(* IEC 61131-3 sources: daoli-st-library/DL_MathData (part 18) *)

(* ---- FC_DL_LrealToFixedField.st ---- *)
(*==============================================================================
 * 组件名称 (Component)  : FC_DL_LrealToFixedField
 * 溯源说明 (Provenance): 道莅 clean-room 防御性实现（IEC 61131-3 纯净实现，闭源文档仅借语义，零代码行）
 * 所属子库 (Sublibrary) : DL_MathData / DataFormat
 * 当前版本 (Version)    : 1.0.0
 * 兼容性   (Platform)   : CODESYS 3.5 / TwinCAT 3 / 汇川 InoProShop / 施耐德
 *                         Machine Expert；纯 IEC 61131-3（第 3 版），仅用
 *                         Standard.library 的 MID / CONCAT / LEN / ABS / TRUNC / LIMIT
 * 组件分类 (Category)   : 函数（FUNCTION）· 纯函数 · 浮点 → 定宽定点文本
 * 功能一句话 (Summary)  : 把 LREAL 按指定整数位宽与小数位数输出成定宽定点文本
 *                         （四舍五入或截断、可选强制正号），非有限输入拒绝输出。
 *
 * 【填充与对齐规则（与 FC_DL_IntToFixedField 共用同一段口径原文）】
 *   ① 右对齐：数值永远贴字段右端，填充字符只在左侧。
 *   ② 本件无 bZeroPad 引脚，整数部分统一用**空格**填充到 uIntDigits 位
 *      ——即 #1 的 bZeroPad = FALSE 分支口径；领先零一律压成空格，
 *      但至少保留一位数字（0.5 输出 "0.500" 而非 ".500"）。
 *   ③ 符号位占一位：**恒留一格**（无符号时填空格），故字段总宽恒为
 *      1 + uIntDigits + (uDecDigits > 0 ? 1 + uDecDigits : 0) ≤ 23，
 *      定长报文的列位由此确定，不随数值正负漂移。
 *   ④ 宽度是契约：uIntDigits / uDecDigits 越界只钳位（0460 信息级）；
 *      整数部分装不下时不截断，直接饱和到全 9 并置 bSaturated。
 *
 * 本件存在的意义 (Why this unit exists)
 *   MES 称重/流量报文要的是「固定小数位、列位对齐」的数值域（"  1234.567"）。
 *   平台内建 LREAL_TO_STRING 的小数位口径与科学计数法门槛三平台不一致
 *   （CODESYS / TwinCAT / InoProShop 对同一值可能给出不同尾数与指数形式），
 *   故本件**禁用** LREAL_TO_STRING，自行按 10 的幂分解：绝对值域取整 → 逐位
 *   分解 → 拼接，末位再加符号，天然对称，输出可在三平台逐字节比对。
 *
 * 边界安全 (Boundary)
 *   ① 非有限输入：NaN 用自不等判据 (x−x) <>(x−x)，±Inf 用 ABS(x) > DBL_MAX
 *      精确判据（R79，禁近似阈值）→ 故障 03AE、bValid = FALSE，
 *      **绝不输出 'NaN' / 'Inf' 冒充合法报文**；
 *   ② uIntDigits 钳 1~15、uDecDigits 钳 0~6，越界钳位 + 信息 0460；
 *   ③ 字段装不下（1 + 整数位 + 1 + 小数位 > 24）→ 故障 03AF。钳位后最大为
 *      23，本分支结构性不可达，属纯防御纵深（R94 统一后处理）；
 *   ④ 整数部分有效位超 uIntDigits → 饱和全 9 + bSaturated + 信息 0461，
 *      bValid 保持 TRUE（饱和可观测，与「非有限」性质不同）；
 *   ⑤ 四舍五入实际进位导致整数位溢出 → 同一饱和路径（复用 0461，不新开码，R90）；
 *   ⑥ 舍入进位未溢出整数位 → 信息 0460 复用（R90 不加码，头注释写明复用理由）；
 *   ⑦ 全部取整只用 TRUNC 作用于**小于 10 的商与小于 10^d 的余数**，绝不 TRUNC
 *      大数，因此任何平台都不会在内建转换上溢出。
 * 遗留假设 (Assumption)
 *   整数部分超过 15 位十进制时 LREAL 已无精确表示（2^53 ≈ 9.007E15），
 *   本件按「输入本身已失真」处理，不承诺末位准确；这也是把
 *   uIntDigits 上限定为 15 的原因（DL_FF_INTMAX）。
 *   逐位分解的商与余数为浮点运算，末位可能受二进制表示误差影响 ±1 个最小
 *   单位（已在四舍五入阈值中吸收），不承诺与十进制手算逐位一致。
 *
 * 错误码    : 16#0001_0460 整数位/小数位已钳位，或四舍五入发生进位——信息级，正常防御
 *             16#0001_0461 整数部分有效位超出字段宽度，已饱和为全 9——信息级，饱和可观测
 *             16#0001_03AE 输入非有限（NaN / ±Inf），拒绝输出——故障级，返回 FALSE
 *             16#0001_03AF 字段宽度装不下（整数位+小数位+符号+小数点超上限）——故障级
 *             16#0001_03B0 预留禁用（故障级，不得挪用）
 * 码位总账  : 16#0001_0460 用 / 16#0001_0461 用 ｜ 16#0001_03AE 用 / 16#0001_03AF 用 / 16#0001_03B0 预留
 * 状态机    : N/A —— 纯函数无顺序状态机
 * 采样约定  : 纯组合函数，无定时器、无内部驻留状态
 * 依赖说明  : 无 DL_ 内部依赖；仅 Standard.library 的 MID / CONCAT / LEN / ABS / TRUNC / LIMIT
 * 验收向量  : V1 1234.5678/整数6/小数3/四舍五入 → '  1234.568'，写 11，TRUE
 *             V2 -42.5/整数6/小数3/截断 → '   -42.500'，写 11，TRUE
 *             V3 0.5/整数2/小数2 → '  0.50'，写 6，TRUE（领先零压成空格但保留一位）
 *             V4 999999.9999/整数6/小数3/四舍五入 → 饱和全 9 ' 999999.999'，
 *                bSaturated=TRUE，eErr=0461，TRUE（进位溢出主向量）
 *             V5 NaN → FALSE，sField=''，eErr=03AE，bError=TRUE
 *             V6 +Inf → FALSE，eErr=03AE
 *             V7 整数位 0 / 小数位 9 → 钳到 1 / 6 且 eErr=0460，仍返回 TRUE
 *             V8 1.0E16/整数15/小数0 → 饱和全 9（失真声明主向量）
 * 红线自检  : 全局变量声明零使用 / 外部变量访问零使用 / 物理地址零使用 ｜ 纯 IEC 61131-3（零厂商转换）
 *             浮点无判等比较（仅自不等 NaN 判据与容差阈值）｜ 除法前置判零
 *             （fPow 恒 ≥ 1.0，构造性非零）｜ 循环全部带守卫 ｜ 数组下标前置界检
 *             全变量双语同行注释 ｜ 状态机 N/A ｜ 无定时器实例 ｜ 无魔法数
 * 修订历史  : 2026-11-16  v1.0.0  首版入库（R22 · 批 1 · 定宽数值字段族）
 *============================================================================*)

FUNCTION FC_DL_LrealToFixedField : BOOL
VAR_INPUT
    fValue      : LREAL;                       // 待编码浮点值，任意有限值 / value to encode, any finite value
    uIntDigits  : UINT := 6;                   // 整数部分最少字符数 [字符]，范围 1~15 / minimum integer characters, range 1~15
    uDecDigits  : UINT := 3;                   // 小数位数 [位]，范围 0~6 / decimal digits, range 0~6
    bRound      : BOOL := TRUE;                // TRUE 四舍五入 / FALSE 向零截断 / TRUE rounds half up, FALSE truncates
    bForceSign  : BOOL := FALSE;               // 正数是否强制 '+' 号 / force '+' sign on positive values
END_VAR
VAR_OUTPUT
    sField      : STRING(24);                  // 定宽定点文本，右对齐 [ASCII] / fixed width fixed point text, right aligned
    uFieldLen   : UINT;                        // 实际写入字符数 [字符] / actual written length [char]
    bSaturated  : BOOL;                        // 整数部分已饱和为全 9 / integer part saturated to all nines
    eErr        : UDINT;                       // 错误码，0 表示无错 / error code, 0 means no error
    bError      : BOOL;                        // 故障级标志，仅故障级错误置位 / fault-class flag, set only on fault-level codes
    bValid      : BOOL;                        // 结果可用标志（饱和时仍为 TRUE） / result usable flag, still TRUE when saturated
END_VAR
VAR
    nIntUse     : INT;                         // 生效整数位宽 [字符]，已钳位 1~15 / effective integer width, clamped
    nDecUse     : INT;                         // 生效小数位数 [位]，已钳位 0~6 / effective decimal digits, clamped
    nTotal      : INT;                         // 字段总宽 [字符] / total field width
    nLead       : INT;                         // 首个非零整数位下标 [索引]，0 表示全零 / index of the first non-zero integer digit, 0 when all zero
    nI          : INT;                         // 通用循环下标 [索引] / general loop index
    nJ          : INT;                         // 升序循环变量（镜像下标用）[索引] / ascending loop var for mirrored index
    nGuard      : INT;                         // 循环守卫计数器 [次] / loop guard counter
    nFracMax    : LINT;                        // 小数位满量 10^nDecUse [无量纲] / full range of the decimal part
    liFrac      : LINT;                        // 小数部分放大后的整数值 [无量纲] / scaled integer value of the decimal part
    liDig       : LINT;                        // 单步取位结果 [无量纲] / single digit extraction result
    bNeg        : BOOL;                        // 输入为负 / input is negative
    bNeedSign   : BOOL;                        // 是否输出符号字符 / whether a sign character is emitted
    bAllNine    : BOOL;                        // 饱和全 9 路径 / saturated all-nines path
    bCarry      : BOOL;                        // 舍入发生进位 / rounding produced a carry
    bPropagate  : BOOL;                        // 进位仍在传播 / the carry is still propagating
    fAbs        : LREAL;                       // 输入绝对值 [无量纲] / absolute value of the input
    fRem        : LREAL;                       // 未分解的剩余量 [无量纲] / remaining undecomposed value
    fPow        : LREAL;                       // 当前位的 10 的幂 [无量纲] / power of ten of the current position
    fIntLimit   : LREAL;                       // 整数部分容量 10^nIntUse [无量纲] / integer capacity
    fFracScaled : LREAL;                       // 放大后的小数部分 [无量纲] / scaled decimal part
    fDiff       : LREAL;                       // NaN 自不等判据的中间量 [无量纲] / intermediate for the NaN self-inequality test
    aInt        : ARRAY[1..15] OF USINT;       // 整数位数字缓存，1 基 [无量纲] / integer digit cache, 1-based
    aDec        : ARRAY[1..6] OF USINT;        // 小数位数字缓存，1 基 [无量纲] / decimal digit cache, 1-based
    sInt        : STRING(15);                  // 整数段（含空格填充）[ASCII] / integer segment including space padding
    sFrac       : STRING(6);                   // 小数段 [ASCII] / decimal segment
    sSign       : STRING(1);                   // 符号段，无符号时填空格 [ASCII] / sign segment, a space when unsigned
    sDigitCh    : STRING(1);                   // 单字符数字，由数字表取出 [ASCII] / single digit character taken from the table
END_VAR
VAR CONSTANT
    DL_FF_MAXLEN   : UINT := 24;               // STRING(24) 物理上限 [字符]，禁写成 255 / physical bound of STRING(24), never 255
    DL_FF_INTMAX   : UINT := 15;               // 整数位宽上限 [字符]，受 2^53 精度约束 / integer width ceiling, bounded by 2^53
    DL_FF_DECMAX   : UINT := 6;                // 小数位数上限 [位] / decimal digit ceiling
    DL_FF_MAXLEN_I : INT := 24;                // 字段上限的 INT 副本 [字符] / INT copy of the field ceiling
    DL_INT_MIN     : INT := 1;                 // 整数位宽下限 [字符] / integer width floor
    DL_DEC_MIN     : INT := 0;                 // 小数位数下限 [位] / decimal digit floor
    DL_INT_MAX     : INT := 15;                // 整数位宽上限的 INT 副本 [字符] / INT copy of the integer width ceiling
    DL_DEC_MAX     : INT := 6;                 // 小数位数上限的 INT 副本 [位] / INT copy of the decimal digit ceiling
    DL_U_ZERO      : UINT := 0;                // 无符号零值 [无量纲] / unsigned zero
    DL_U_ONE       : UINT := 1;                // 无符号一值 [无量纲] / unsigned one
    DL_ONE_I       : INT := 1;                 // 整型一，用于 FOR 起始 [无量纲] / integer one used as a FOR start
    DL_SIGN_RES    : INT := 1;                 // 符号位恒留宽度 [字符] / reserved sign position width
    DL_POINT_W     : INT := 1;                 // 小数点占位宽度 [字符] / decimal point width
    DL_DIG_LAST    : INT := 9;                 // 单个数字位最大值 [无量纲] / maximum single digit value
    DL_GUARD_MAX   : INT := 20;                // 循环守卫上限 [次] / loop guard ceiling
    DL_TEN_I       : INT := 10;                // 十进制基数的 INT 副本 [无量纲] / INT copy of the decimal radix
    DL_TEN_L       : LINT := 10;               // 十进制基数的 LINT 副本 [无量纲] / LINT copy of the decimal radix
    DL_TEN_R       : LREAL := 10.0;            // 十进制基数的 LREAL 副本 [无量纲] / LREAL copy of the decimal radix
    DL_ONE_R       : LREAL := 1.0;             // 实型一，幂循环起点 [无量纲] / real one, power loop start
    DL_HALF_R      : LREAL := 0.5;             // 四舍五入偏置 [无量纲] / half-up rounding offset
    DL_LREAL_MAX   : LREAL := 1.7976931348623157E308; // LREAL 最大有限值，±Inf 精确判据 / maximum finite LREAL, exact infinity test
    DL_DIGITS      : STRING(10) := '0123456789'; // 数字字符表，经 MID 取值 [ASCII] / digit table read through MID
    DL_POINT_CH    : STRING(1) := '.';         // 小数点字符 [字符] / decimal point character
    DL_SPACE_CH    : STRING(1) := ' ';         // 空格填充字符 [字符] / space pad character
    DL_SIGN_PLUS   : STRING(1) := '+';         // 正号字符 [字符] / plus sign character
    DL_SIGN_MINUS  : STRING(1) := '-';         // 负号字符 [字符] / minus sign character
    DL_CH_ONE      : INT := 1;                 // MID 的单字符长度 [字符] / single character length for MID
END_VAR

(*------------------------------------------------------------------------------
 * 段 1｜返回值与输出预置（L1/L9：任何早退路径不留脏值）
 *      Preset the return value and every output, no stale value on any exit
 *-----------------------------------------------------------------------------*)
FC_DL_LrealToFixedField := FALSE;              // 返回值预置失败 / preset to FALSE
sField      := '';                             // 字段清空 / field cleared
uFieldLen   := 0;                              // 写入长度预置 0 [字符] / written length preset to zero
bSaturated  := FALSE;                          // 饱和标志预置 FALSE / saturation preset to FALSE
eErr        := 16#0000_0000;                   // 错误码预置无错 / error code preset to none
bError      := FALSE;                          // 故障标志预置 FALSE / fault flag preset to FALSE
bValid      := FALSE;                          // 结果可用预置 FALSE / usable flag preset to FALSE
nIntUse     := DL_INT_MIN;                     // 整数位宽预置下限 / integer width preset to the floor
nDecUse     := DL_DEC_MIN;                     // 小数位数预置下限 / decimal digits preset to the floor
nTotal      := 0;                              // 总宽预置 0 / total width preset to zero
nLead       := 0;                              // 领先零位置预置 0 / leading position preset to zero
nGuard      := 0;                              // 守卫预置 0 / guard preset to zero
nFracMax    := 1;                              // 小数满量预置 1 / decimal full range preset to one
liFrac      := 0;                              // 小数整数化预置 0 / scaled decimal preset to zero
liDig       := 0;                              // 取位结果预置 0 / digit result preset to zero
bNeg        := FALSE;                          // 负号标志预置 FALSE / negative flag preset to FALSE
bNeedSign   := FALSE;                          // 符号标志预置 FALSE / sign flag preset to FALSE
bAllNine    := FALSE;                          // 饱和路径预置 FALSE / saturation path preset to FALSE
bCarry      := FALSE;                          // 进位标志预置 FALSE / carry flag preset to FALSE
bPropagate  := FALSE;                          // 进位传播预置 FALSE / propagation preset to FALSE
fAbs        := 0.0;                            // 绝对值预置 0 / absolute value preset to zero
fRem        := 0.0;                            // 剩余量预置 0 / remainder preset to zero
fPow        := DL_ONE_R;                       // 幂预置 1 / power preset to one
fIntLimit   := DL_ONE_R;                       // 整数容量预置 1 / integer capacity preset to one
fFracScaled := 0.0;                            // 放大值预置 0 / scaled value preset to zero
sSign       := DL_SPACE_CH;                    // 符号段预置空格（符号位恒留一格） / sign segment preset to a space, the position is always reserved

(*------------------------------------------------------------------------------
 * 段 2｜非有限输入闸门（R79 精确判据：NaN 自不等 + ±Inf 与 DBL_MAX 直比）
 *      Non-finite gate with exact criteria, no approximate thresholds
 *-----------------------------------------------------------------------------*)
fDiff := fValue - fValue;                      // 有限值得 0，NaN 得 NaN / zero for finite input, NaN for NaN input
IF fDiff <> fDiff THEN
    eErr   := 16#0001_03AE;                    // 故障级：NaN 输入 / fault: NaN input
    bError := TRUE;                            // 置故障标志 / raise the fault flag
    bValid := FALSE;                           // 结果不可用 / result unusable
    sField := '';                              // 绝不输出 'NaN' 冒充合法报文 / never emit NaN as a legal field
    RETURN;                                    // 早退路径已统一后处理 / the early exit is fully post-processed
END_IF
IF ABS(fValue) > DL_LREAL_MAX THEN
    eErr   := 16#0001_03AE;                    // 故障级：±Inf 输入 / fault: infinity input
    bError := TRUE;                            // 置故障标志 / raise the fault flag
    bValid := FALSE;                           // 结果不可用 / result unusable
    sField := '';                              // 绝不输出 'Inf' 冒充合法报文 / never emit Inf as a legal field
    RETURN;
END_IF

(*------------------------------------------------------------------------------
 * 段 3｜位宽钳位（越界只钳位；信息级码不置 bError）
 *      Width clamping, out-of-range values are clamped and never raise bError
 *-----------------------------------------------------------------------------*)
IF uIntDigits < DL_U_ONE THEN
    nIntUse := DL_INT_MIN;                     // 钳到下限 1 / clamped to the floor
    eErr    := 16#0001_0460;                   // 信息级：整数位已钳位 / informational: integer width clamped
ELSIF uIntDigits > DL_FF_INTMAX THEN
    nIntUse := DL_INT_MAX;                     // 钳到上限 15 / clamped to the ceiling
    eErr    := 16#0001_0460;                   // 信息级：整数位已钳位 / informational: integer width clamped
ELSE
    nIntUse := UINT_TO_INT(uIntDigits);         // 域内直通 / passed through inside the domain
END_IF

IF uDecDigits > DL_FF_DECMAX THEN
    nDecUse := DL_DEC_MAX;                     // 钳到上限 6 / clamped to the ceiling
    eErr    := 16#0001_0460;                   // 信息级：小数位已钳位 / informational: decimal digits clamped
ELSE
    nDecUse := UINT_TO_INT(uDecDigits);         // 域内直通（无符号量无下限问题） / passed through, no floor issue for unsigned
END_IF

(*------------------------------------------------------------------------------
 * 段 4｜字段容量闸门（防御纵深：钳位后最大 23，本分支结构性不可达）
 *      Capacity gate, structurally unreachable after clamping, pure defense in depth
 *-----------------------------------------------------------------------------*)
nTotal := DL_SIGN_RES + nIntUse;                // 符号位恒留一格 + 整数位 / reserved sign plus integer width
IF nDecUse > DL_DEC_MIN THEN
    nTotal := nTotal + DL_POINT_W + nDecUse;    // 有小数位时加小数点与小数位 / add the point and the decimal digits
END_IF
IF nTotal > DL_FF_MAXLEN_I THEN
    eErr   := 16#0001_03AF;                     // 故障级：字段装不下 / fault: the field cannot hold the value
    bError := TRUE;                             // 置故障标志 / raise the fault flag
    bValid := FALSE;                            // 结果不可用 / result unusable
    sField := '';                               // 字段保持空串 / field stays empty
    RETURN;
END_IF

(*------------------------------------------------------------------------------
 * 段 5｜符号判定、整数量级与饱和预判（先判容量，绝不 TRUNC 大数）
 *      Sign, integer magnitude and saturation pre-check, never TRUNC a large value
 *-----------------------------------------------------------------------------*)
bNeg      := (fValue < 0.0);                    // 负值判据 / negative test
bNeedSign := bNeg OR bForceSign;                // 负号必需，正号由引脚决定 / minus always needed, plus only when forced
IF bNeedSign THEN
    IF bNeg THEN
        sSign := DL_SIGN_MINUS;                 // 负号 / minus sign
    ELSE
        sSign := DL_SIGN_PLUS;                  // 强制正号 / forced plus sign
    END_IF
ELSE
    sSign := DL_SPACE_CH;                       // 无符号：占位填空格，保持字段恒宽 / unsigned, a space keeps the width constant
END_IF

fAbs := ABS(fValue);                            // 绝对值域运算，末位再加符号，正负对称 / absolute domain, the sign is added at the end
fIntLimit := DL_ONE_R;                          // 容量初值 1 / capacity starts at one
FOR nI := DL_ONE_I TO nIntUse DO
    fIntLimit := fIntLimit * DL_TEN_R;          // 容量 = 10^nIntUse，nIntUse ≤ 15 在 LREAL 精确域内 / capacity, exact for n <= 15
END_FOR
IF fAbs >= fIntLimit THEN
    bAllNine := TRUE;                           // 整数部分装不下：饱和全 9，不进分解 / overflow, saturate to all nines
    eErr     := 16#0001_0461;                   // 信息级：整数部分已饱和 / informational: integer part saturated
    bSaturated := TRUE;                         // 饱和可观测 / saturation observable
END_IF

(*------------------------------------------------------------------------------
 * 段 6｜整数位逐位分解（TRUNC 只作用于小于 10 的商）
 *      Integer digit decomposition, TRUNC only ever sees a quotient below ten
 *-----------------------------------------------------------------------------*)
IF NOT bAllNine THEN
    fRem := fAbs;                               // 从绝对值开始分解 / decomposition starts from the absolute value
    fPow := DL_ONE_R;                           // 最高位幂初值 1 / highest power starts at one
    FOR nI := DL_ONE_I TO (nIntUse - DL_ONE_I) DO
        fPow := fPow * DL_TEN_R;                // 幂升到 10^(nIntUse-1) / raise to the highest power
    END_FOR
    FOR nI := DL_ONE_I TO nIntUse DO
        IF fPow > 0.0 THEN
            liDig := TRUNC(fRem / fPow);        // 商恒 0~9，TRUNC 永不溢出 / quotient always 0~9, TRUNC never overflows
        ELSE
            liDig := 0;                         // 构造性不可达的兜底 / structurally unreachable fallback
        END_IF
        IF liDig < 0 THEN
            liDig := 0;                         // 下界夹紧 / clamped low
        ELSIF liDig > DL_DIG_LAST THEN
            liDig := DL_DIG_LAST;               // 上界夹紧 / clamped high
        END_IF
        aInt[nI] := LINT_TO_USINT(liDig);       // 缓存本位数 / cache this digit
        fRem := fRem - LINT_TO_LREAL(liDig) * fPow; // 扣掉已分解部分 / subtract the decomposed part
        fPow := fPow / DL_TEN_R;                // 幂降一位 / step down one power
    END_FOR
    IF fRem < 0.0 THEN
        fRem := 0.0;                            // 浮点误差兜底，剩余量恒非负 / floating point fallback, the remainder stays non-negative
    END_IF

    (* 小数部分：放大到整数域后取整，四舍五入加 0.5（负值已处理成绝对值，天然对称） *)
    (* Decimal part, scaled to the integer domain, half-up adds 0.5 in the absolute domain *)
    nFracMax := 1;                              // 小数满量初值 1 / full range starts at one
    FOR nI := DL_ONE_I TO nDecUse DO
        nFracMax := nFracMax * DL_TEN_L;        // 满量 = 10^nDecUse，nDecUse ≤ 6 / full range, n <= 6
    END_FOR
    fFracScaled := fRem * LINT_TO_LREAL(nFracMax);// 放大到小数满量 [无量纲] / scaled up to the decimal range
    IF bRound THEN
        fFracScaled := fFracScaled + DL_HALF_R;  // 四舍五入偏置 / half-up offset
    END_IF
    liFrac := TRUNC(fFracScaled);                // 取值恒 ≤ 10^nDecUse < 1.0E7，TRUNC 安全 / always below 1E7, TRUNC is safe
    IF liFrac < 0 THEN
        liFrac := 0;                             // 下界夹紧 / clamped low
    END_IF
    IF liFrac >= nFracMax THEN
        liFrac := liFrac - nFracMax;             // 满量即归零 / wrapped to zero
        bCarry := TRUE;                          // 向整数位进位 / carry into the integer part
    END_IF

    (* 进位传播：从最低整数位向前逐位加一，全 9 则整体饱和 *)
    (* Carry propagation from the least significant integer digit, all nines saturate everything *)
    IF bCarry THEN
        eErr        := 16#0001_0460;             // 信息级：舍入进位（复用 0460，R90 不加码） / informational: rounding carried, code reused
        nLead       := nIntUse;                  // 传播从最低位开始 / propagation starts at the lowest digit
        bPropagate  := TRUE;                     // 传播仍在进行 / the carry is still propagating
        nGuard      := 0;                        // 守卫清零 / guard cleared
        WHILE bPropagate AND (nLead >= DL_ONE_I) AND (nGuard <= DL_GUARD_MAX) DO
            IF aInt[nLead] < DL_DIG_LAST THEN
                aInt[nLead] := aInt[nLead] + 1;  // 本位加一，传播结束 / increment and stop propagating
                bPropagate  := FALSE;
            ELSE
                aInt[nLead] := 0;                // 本位满 9 归零，继续向前 / wrap to zero and keep propagating
                nLead := nLead - DL_ONE_I;
            END_IF
            nGuard := nGuard + DL_ONE_I;         // 守卫累计 / guard incremented
        END_WHILE
        IF bPropagate THEN
            bAllNine := TRUE;                    // 整数位全部溢出：饱和全 9 / every integer digit overflowed
            eErr     := 16#0001_0461;            // 信息级：整数部分已饱和 / informational: integer part saturated
            bSaturated := TRUE;                  // 饱和可观测 / saturation observable
        END_IF
    END_IF
END_IF

(*------------------------------------------------------------------------------
 * 段 7｜饱和路径填 9（整数位与小数位同时置 9，语义为「超出可表示范围」）
 *      Saturation path fills nines, meaning the value exceeds the representable range
 *-----------------------------------------------------------------------------*)
IF bAllNine THEN
    FOR nI := DL_ONE_I TO nIntUse DO
        aInt[nI] := INT_TO_USINT(DL_DIG_LAST);   // 整数位全 9 / integer digits all nine
    END_FOR
    FOR nI := DL_ONE_I TO nDecUse DO
        aDec[nI] := INT_TO_USINT(DL_DIG_LAST);   // 小数位全 9 / decimal digits all nine
    END_FOR
    liFrac := 0;                                 // 小数整数化量不再使用 / the scaled decimal value is no longer used
ELSE
    (* 小数位逐位分解：从小到大取余，负域无需用（值恒非负） *)
    (* Decimal digit decomposition, the value is always non-negative here *)
    FOR nJ := DL_ONE_I TO nDecUse DO
        nI := nDecUse - nJ + DL_ONE_I;       // 镜像下标：R509 禁 DOWNTO / mirrored index, DOWNTO unsupported
        aDec[nI] := LINT_TO_USINT(liFrac MOD DL_TEN_L); // 取最低位 / take the least significant digit
        liFrac   := liFrac / DL_TEN_L;           // 降一位 / step down
    END_FOR
END_IF

(*------------------------------------------------------------------------------
 * 段 8｜领先零定位（压成空格，但至少保留一位数字）
 *      Locate the leading zeros, replaced by spaces while keeping at least one digit
 *-----------------------------------------------------------------------------*)
nLead := 0;                                      // 0 表示尚未找到非零位 / zero means no non-zero digit found yet
FOR nI := DL_ONE_I TO nIntUse DO
    IF (nLead = 0) AND (aInt[nI] <> 0) THEN
        nLead := nI;                             // 记录首个非零位 / remember the first non-zero position
    END_IF
END_FOR
IF nLead = 0 THEN
    nLead := nIntUse;                            // 全零：最后一位仍输出 '0' / all zero, the last position still prints a zero
END_IF

(*------------------------------------------------------------------------------
 * 段 9｜拼装（整数段 + 小数点 + 小数段，符号段恒占一格）
 *      Assembly, integer segment plus point plus decimals, the sign position is always reserved
 *-----------------------------------------------------------------------------*)
sInt := '';                                      // 整数段清空 / integer segment cleared
FOR nI := DL_ONE_I TO nIntUse DO
    IF nI < nLead THEN
        sInt := CONCAT(sInt, DL_SPACE_CH);        // 领先零压成空格 / a leading zero becomes a space
    ELSE
        sDigitCh := MID(DL_DIGITS, DL_CH_ONE, USINT_TO_INT(aInt[nI]) + DL_CH_ONE); // 数字 → 字符（查表） / digit to character by table
        sInt := CONCAT(sInt, sDigitCh);           // 追加数字 / append the digit
    END_IF
END_FOR

sFrac := '';                                     // 小数段清空 / decimal segment cleared
FOR nI := DL_ONE_I TO nDecUse DO
    sDigitCh := MID(DL_DIGITS, DL_CH_ONE, USINT_TO_INT(aDec[nI]) + DL_CH_ONE); // 数字 → 字符（查表） / digit to character by table
    sFrac := CONCAT(sFrac, sDigitCh);             // 追加小数位 / append the decimal digit
END_FOR

sField := CONCAT(sSign, sInt);                   // 符号位 + 整数段 / sign position plus integer segment
IF nDecUse > DL_DEC_MIN THEN
    sField := CONCAT(sField, DL_POINT_CH);        // 小数点 / decimal point
    sField := CONCAT(sField, sFrac);              // 小数段 / decimal segment
END_IF

(*------------------------------------------------------------------------------
 * 段 10｜长度复检与出口（结构性不可达，纯防御纵深）
 *      Length recheck and exit, structurally unreachable, pure defense in depth
 *-----------------------------------------------------------------------------*)
IF LEN(sField) <> nTotal THEN
    eErr   := 16#0001_03AF;                       // 复检不符：按字段容量故障处理 / recheck mismatch, capacity fault
    bError := TRUE;                               // 置故障标志 / raise the fault flag
    bValid := FALSE;                              // 结果不可用 / result unusable
    sField := '';                                 // 字段回空，绝不交出不完整字段 / field emptied
    uFieldLen := 0;                               // 写入长度回 0 / written length back to zero
    RETURN;
END_IF

uFieldLen := INT_TO_UINT(nTotal);                  // 写入字符数 = 设计总宽 / written length equals the designed width
bValid    := TRUE;                                 // 结果可用（饱和亦为可用，降级可观测） / usable even when saturated
FC_DL_LrealToFixedField := TRUE;                   // 编码成功 / encoding succeeded
END_FUNCTION

(* ---- FC_DL_LrealToLintSat.st ---- *)
(*
    FC_DL_LrealToLintSat —— LREAL 到 LINT 域外饱和转换
    ------------------------------------------------------------------
    分类      : DL_MathData / Convert
    前缀      : FC_DL_
    版本      : 1.0.0
    溯源      : IEC 61131-3 标准语义的道莅防御性实现
                （接口语义由 IEC 61131-3 定义，内部委托平台内建 TRUNC 与 LREAL_TO_LINT，
                  外围统一错误码 / 钳位 / 双语文档；clean-room 重写，
                  未复制任何闭源厂商源码，参考实现仅限 MIT/Apache 许可）
    平台      : 纯 IEC 61131-3，CODESYS / TwinCAT / InoProShop 通用
    作者      : 道莅代码库 · PLC编程专家（R17）
    ------------------------------------------------------------------
    功能说明  : 将 LREAL 防御性转换为 LINT 并作为返回值输出；
                非有限输入（NaN 或 ±INF）判为故障级 16#0001_02F4，返回 0 且 bValid=FALSE；
                取整取向声明：向零截断（TRUNC 语义）后钳位，与 FC_DL_RealToLintSat 及
                R16 FC_DL_LrealToDintSat 同口径；
                与 FC_DL_RealToLintSat 的职责边界：源类型不同（IEC 61131-3 无 ANY_REAL 泛型），
                双版本是库内既定策略（R16 饱和转换族先例），不做类型合并；
                域外按方向饱和（上界 9223372036854775807 / 下界负向极值）
                并置信息级 16#0001_0230；下界用 -DL_LINT_MAX - 1 计算式，禁负数字面量直写；
                钳位方向：双侧饱和，绝不回绕。
    错误码    : 16#0001_0230 输入超 LINT 域，已按符号饱和——信息级，正常防御
                16#0001_0231 预留禁用（信息级，不得挪用）
                16#0001_02F4 非有限输入（NaN 或 ±INF）——故障级，返回 0
                16#0001_02F5 预留禁用（故障级，不得挪用）
                16#0001_02F6 预留禁用（故障级，不得挪用）
    状态机    : R6 标注 N/A —— 本组件为纯函数无顺序状态机，无 CASE 可写，非法状态不可能出现，故以本节说明替代 ELSE 兜底
    修订记录  : 2026-11-16 v1.0.0 首次入库（R17）
*)
FUNCTION FC_DL_LrealToLintSat : LINT
VAR_INPUT
    fIn : LREAL; // 待转换 64 位浮点值，建议域 ±9.2E18（非有限拦截，域外饱和） [无量纲] / 64-bit floating value to convert, suggested domain +/-9.2E18 [dimensionless]
END_VAR
VAR_OUTPUT
    eErr   : UDINT; // 错误码，0=正常 / error id, 0=ok
    bError : BOOL;  // 是否出错，eErr 非 0 时为 TRUE / error flag, TRUE when eErr is nonzero
    bValid : BOOL;  // 输出是否有效可用 / output valid flag
END_VAR
VAR CONSTANT
    DL_LINT_MAX_LR    : LREAL := 9.2233720368547758E18;          // LINT 域上界在 LREAL 域的精确可表近似值 [无量纲] / LINT upper bound represented in LREAL [dimensionless]
    DL_LINT_MAX       : LINT  := 9223372036854775807;            // LINT 上界饱和输出值 [无量纲] / LINT upper saturation output [dimensionless]
    DL_LINT_ZERO      : LINT  := 0;                              // 故障缺省返回值 [无量纲] / fault default return value [dimensionless]
    DL_LREAL_HUGE     : LREAL := 1.7976931348623157E308;         // LREAL 最大有限幅值，超过即判 ±INF [无量纲] / max finite LREAL magnitude, beyond means +/-INF [dimensionless]
END_VAR
VAR
    bNonFinite : BOOL; // 非有限（NaN 或 ±INF）判定结果 / non-finite (NaN or +/-INF) detection result
END_VAR

// 段 1｜返回值与错误状态预置 / segment 1, preset return value and error status
FC_DL_LrealToLintSat := DL_LINT_ZERO; // 故障缺省返回 0 [无量纲] / fault default 0 [dimensionless]
eErr   := 0;     // 预置无错误 / preset no error
bError := FALSE; // 预置无故障 / preset no fault
bValid := FALSE; // 预置输出无效，通过三路闸后置位 / preset invalid, set TRUE after the three gates

// 段 2｜非有限防御闸 / segment 2, non-finite guard
bNonFinite := (fIn <> fIn) OR (fIn > DL_LREAL_HUGE) OR (fIn < -DL_LREAL_HUGE); // 非有限判定（NaN 自不等 + 最大有限幅值判 ±INF） [无量纲] / non-finite check (NaN by self-inequality, +/-INF by max finite magnitude) [dimensionless]
IF bNonFinite THEN
    eErr := 16#0001_02F4; // 非有限输入故障码 / non-finite input fault id
    bError := TRUE;       // 置故障标志 / raise error flag
    bValid := FALSE;      // 输出不可用 / output not usable
    RETURN;               // 故障级提前返回，保持缺省 0 / early return on fault, keep default 0
END_IF

// 段 3｜域外判定饱和与域内截断转换（末段） / segment 3, out-of-domain saturation and in-domain truncate conversion (final)
IF fIn > DL_LINT_MAX_LR THEN
    FC_DL_LrealToLintSat := DL_LINT_MAX; // 上界饱和至 LINT 上界 [无量纲] / saturate to the LINT upper bound [dimensionless]
    eErr := 16#0001_0230;                // 信息级：域外饱和，正常防御 / info level: out-of-domain saturation, normal defence
    bError := FALSE;                     // 信息级不置故障 / info level never raises fault
    bValid := TRUE;                      // 饱和值本身有效可用 / the saturated value itself is valid
    RETURN;                              // 饱和即出口 / saturation is the exit
ELSIF fIn < -DL_LINT_MAX_LR THEN
    FC_DL_LrealToLintSat := -DL_LINT_MAX - 1; // 下界饱和，用计算式书写，等于 LINT 最小值 [无量纲] / saturate to the LINT minimum, written as a computed expression [dimensionless]
    eErr := 16#0001_0230;                     // 上下共用同一业务语义码，方向写进头注释 / both directions share one business-semantics code, directions documented in the header
    bError := FALSE;                          // 信息级不置故障 / info level never raises fault
    bValid := TRUE;                           // 饱和值本身有效可用 / the saturated value itself is valid
    RETURN;                                   // 饱和即出口 / saturation is the exit
ELSE
    FC_DL_LrealToLintSat := LREAL_TO_LINT(TRUNC(fIn)); // 先 TRUNC 成整值再转，取向恒为向零截断 [无量纲] / TRUNC to an integral value before converting, always truncates toward zero [dimensionless]
    eErr := 0;                                         // 域内无错误 / in-domain, no error
END_IF
bError := FALSE; // 信息级不置故障 / info level never raises fault
bValid := TRUE;  // 域内或饱和输出均有效可用 / in-domain or saturated output is valid
END_FUNCTION

(* ---- FC_DL_LrealToRealSat.st ---- *)
(*
    FC_DL_LrealToRealSat —— LREAL 到 REAL 定长饱和防御转换
    ------------------------------------------------------------------
    分类      : DL_MathData / Convert
    前缀      : FC_DL_
    版本      : 1.0.0
    溯源      : IEC 61131-3 标准语义的道莅防御性实现
                （内部委托平台内建函数，外围统一错误码/钳位/双语文档；
                  未复制任何闭源厂商源码，参考实现仅限 MIT/Apache 许可）
    平台      : 纯 IEC 61131-3，CODESYS / TwinCAT / InoProShop 通用
    作者      : 道莅代码库 · PLC编程专家（R16）
    ------------------------------------------------------------------
    功能说明  : 将 LREAL 输入防御性转换为 REAL 并作为返回值输出；
                非有限输入（NaN 或 ±INF）判为故障级 16#0001_028E，返回 0.0 且 bValid=FALSE；
                幅值 |fIn| 超出 REAL 上限 3.402823E38 时按符号双侧饱和钳位，置信息级 16#0001_01C0；
                钳位方向：正向钳至上界 +3.402823E38，负向钳至下界 -3.402823E38（双侧饱和）；
                ±INF 采用平台安全幅值比较判定（阈值取 LREAL 最大有限幅值），NaN 用 fIn <> fIn 自不等判定；
                域内转换委托平台内建 LREAL_TO_REAL 语义，不重实现数学内核；
                信息级码属正常防御：bError=FALSE、bValid=TRUE，输出钳位后防御值。
    错误码    : 16#0001_028E 非有限输入（NaN 或 ±INF）——故障级，返回 0.0
                16#0001_01C0 幅值超 REAL 域，已按符号饱和钳位——信息级，正常防御
                16#0001_01C1 预留禁用（信息级，不得挪用）
                16#0001_028F 预留禁用（故障级，不得挪用）
                16#0001_0290 预留禁用（故障级，不得挪用）
    状态机    : R6 标注 N/A —— 本组件为纯函数无顺序状态机，无 CASE 可写，非法状态不可能出现，故以本节说明替代 ELSE 兜底
    修订记录  : 2026-11-16 v1.0.0 首次入库（R16）
*)
FUNCTION FC_DL_LrealToRealSat : REAL
VAR_INPUT
    fIn : LREAL; // 待转换输入 [无量纲] / input value to convert
END_VAR
VAR_OUTPUT
    eErr   : UDINT; // 错误码，0=正常 / error id, 0=ok
    bError : BOOL;  // 是否出错，eErr 非 0 时为 TRUE / error flag, TRUE when eErr is nonzero
    bValid : BOOL;  // 输出是否有效可用 / output valid flag
END_VAR
VAR CONSTANT
    DL_REAL_MAX   : LREAL := 3.402823E38;            // REAL 域最大有限幅值 [无量纲] / maximum finite magnitude of REAL domain
    DL_LREAL_HUGE : LREAL := 1.7976931348623157E308; // LREAL 最大有限幅值，超过即判 ±INF [无量纲] / max finite LREAL magnitude, beyond means +/-INF
END_VAR
VAR
    bNonFinite : BOOL; // 非有限（NaN 或 ±INF）判定结果 / non-finite (NaN or +/-INF) detection result
END_VAR

// 段 1｜返回值与错误状态预置 / segment 1, preset return value and error status
FC_DL_LrealToRealSat := 0.0; // 故障缺省返回 0 [无量纲] / fault default returns 0
eErr   := 0;     // 预置无错误 / preset no error
bError := FALSE; // 预置无故障 / preset no fault
bValid := FALSE; // 预置无效，通过防御闸后置位 / preset invalid, set TRUE after guard passes

// 段 2｜非有限防御闸 / segment 2, non-finite guard
bNonFinite := (fIn <> fIn) OR (fIn > DL_LREAL_HUGE) OR (fIn < -DL_LREAL_HUGE); // NaN 自不等判定，±INF 用安全幅值比较 [无量纲] / NaN by self-inequality, +/-INF by safe magnitude compare
IF bNonFinite THEN
    FC_DL_LrealToRealSat := 0.0; // 故障级返回 0 [无量纲] / fault level returns 0
    eErr   := 16#0001_028E;      // 非有限输入故障码 / non-finite input fault id
    bError := TRUE;              // 置故障标志 / set fault flag
    bValid := FALSE;             // 输出无效 / output invalid
    RETURN;                      // 立即返回 / immediate return
END_IF

// 段 3｜饱和钳位与主体转换（末段） / segment 3, saturating clamp and main conversion (final)
IF fIn > DL_REAL_MAX THEN
    FC_DL_LrealToRealSat := DL_REAL_MAX; // 正向饱和钳至 REAL 上界 [无量纲] / saturate to REAL upper bound
    eErr := 16#0001_01C0;                // 信息级：超上界已钳位 / info level: above upper bound, clamped
ELSIF fIn < -DL_REAL_MAX THEN
    FC_DL_LrealToRealSat := -DL_REAL_MAX; // 负向饱和钳至 REAL 下界 [无量纲] / saturate to REAL lower bound
    eErr := 16#0001_01C0;                 // 信息级：超下界已钳位 / info level: below lower bound, clamped
ELSE
    FC_DL_LrealToRealSat := LREAL_TO_REAL(fIn); // 域内委托平台内建 _TO_ 转换语义 / in-domain delegate to built-in _TO_ conversion
    eErr := 0; // 域内无错误 / in-domain, no error
END_IF
bError := FALSE; // 信息级钳位不置故障，故障分支已提前返回 / info-level clamp never raises fault, fault branch has returned
bValid := TRUE;  // 域内或钳位输出均有效可用 / in-domain or clamped output is valid
END_FUNCTION

(* ---- FC_DL_LrealToStringTrim.st ---- *)
(*
    FC_DL_LrealToStringTrim —— LREAL 到 STRING 的防御字符串化（非有限值统一文本）
    ------------------------------------------------------------------
    分类      : DL_MathData / Convert
    前缀      : FC_DL_
    版本      : 1.0.1
    溯源      : IEC 61131-3 标准语义的道莅防御性实现（LREAL → STRING，非有限值统一文本）；
                委托平台内建 LREAL_TO_STRING 与标准串函数 LEN / MID / LEFT，本件不重实现格式化内核；
                非有限值判据与统一文本、空格修剪、四步截断样板、错误分级与码位 100% 自有；
                clean-room 重写，未复制任何闭源厂商源码，参考实现仅限 MIT/Apache 许可
    平台      : 纯 IEC 61131-3，CODESYS V3.5+ / TwinCAT 3 / InoProShop 通用
    作者      : 道莅代码库 · PLC编程专家（R20）
    ------------------------------------------------------------------
    功能说明  : 趋势记录、报警文本、报表导出都要把模拟量序列化成文本。有限值的宽度与小数位
                各平台本就不一，非有限值更糟：NaN 在有的平台是 'NaN'，有的是 '1.#QNAN'，
                ±Inf 有 'INF' / 'Infinity' / '1.#INF' / 乱码多种结果，上位机按字符串比对必然漏判。
                核心防御：① 非有限值不走内建转换，直接映射成本库统一的三个字面量
                   'NaN' / 'Inf+' / 'Inf-'：统一文本是可用输出而非故障，故发信息级、
                   bValid 仍为 TRUE——把 NaN 判成故障级会让一个采样坏点牵动整条报警链；
                ② NaN 判定用自反性（x <> x），Inf 判定用「x−x 产 NaN」精确判据 + LREAL
                   最大值幅值兜底，两判据分开置位：
                   IEEE 754 里 NaN 与任何值（含自身）比较均为假，任何容差比较对 NaN 恒假，
                   只能用自反性判据——这是本库浮点判等「一律用 ABS 容差」规则的唯一例外，
                   其余浮点比较（如符号判定）均不做判等；
                   无穷判据同源：任何有限值 x−x 恒为 0（0 <> 0 为假），无穷处 x−x 产 NaN
                   （NaN <> NaN 为真）。R20 终审修正：原判据用幅值阈值 1.79E308，该值落在
                   LREAL 可表域内，会把 [1.79E308, LREAL 最大值] 的合法有限值误判成无穷；
                   现改双判据，幅值兜底阈值提到 LREAL 最大值，残余仅剩「恰为最大值」单值；
                ③ 有限值走内建 + 空格修剪 + 四步截断样板（R37），与整型件同一口径；
                ④ 目标长度 0 结构性钳到 1 字符：零长度目标无意义，
                   钳位后必然触发截断分支，事件由 bTruncated 与信息码体现，不静默。
                职责边界：DINT 字符串化归 FC_DL_DintToStringTrim；字符串转回数值归
                FC_DL_StringToLReal；本件只管 LREAL 方向。
    编译门槛  : 主路径依赖平台内建 LREAL_TO_STRING 与标准串函数 LEN / MID / LEFT。
                LREAL_TO_STRING 的有效位数与宽度平台间不同，故本件不假设宽度，
                一律 LEN 实测后按目标长度钳位；幅值兜底阈值取 LREAL 最大值
                1.7976931348623157E308（不是 1.79E308——后者在 LREAL 域内，会把
                极大有限值误判为无穷，R20 终审修正）。
    错误码    : 16#0001_0428 非有限值已映射统一文本（bNonFinite 可查）——信息级，值可用
                16#0001_0429 发生空格修剪或截断——信息级，值可用
                16#0001_035A 需要截断但 bAllowTrunc = FALSE——故障级，返回空串
                16#0001_035B 预留（故障级，不得挪用）
                16#0001_035C 预留禁用（故障级，不得挪用）
    码位总账  : 16#0001_0428 用 / 16#0001_0429 用 ｜ 16#0001_035A 用 / 16#0001_035B 预留 / 16#0001_035C 预留
    状态机    : R6 标注 N/A —— 本组件为纯函数无顺序状态机，无 CASE 可写，非法状态不可能出现
    采样约定  : 本件无定时器、无沿检测、无状态；单拍纯计算，结论与任务周期无关。
    修订记录  : 2026-11-16 v1.0.0 首次入库（R20）
                2026-11-16 v1.0.1 R20 终审修正：无穷幅值判据阈值由 1.79E308 改为 LREAL 最大值
                 并补 x−x 精确判据，消除极大有限值被误判为 'Inf+' 的缺陷；对外引脚零变更
*)
FUNCTION FC_DL_LrealToStringTrim : STRING(255)
VAR_INPUT
    fIn              : LREAL;                 // 待字符串化的数值 [无量纲]，全域（含 NaN 与 ±Inf）/ value to serialise [dimensionless], full domain including NaN and infinities
    uTargetMax       : USINT := 31;           // 目标缓冲可用长度 [字符]，1~255 / usable target length [characters], 1 to 255
    bAllowTrunc      : BOOL := FALSE;         // TRUE = 允许截断；FALSE = 需截断即故障 / TRUE allows truncation, FALSE turns it into a fault
END_VAR
VAR_OUTPUT
    eErr             : UDINT;                 // 错误码，0=正常 / error id, 0=ok
    bError           : BOOL;                  // 故障标志，eErr 为故障级时 TRUE / error flag, TRUE on fault-level eErr
    bValid           : BOOL;                  // 返回值是否可用（故障级为 FALSE）/ return usable, FALSE on fault level
    bNonFinite       : BOOL;                  // 输入为非有限值（NaN 或 ±Inf）/ the input is non-finite, NaN or an infinity
    bTrimmed         : BOOL;                  // 修剪了前导空格 / leading blanks were trimmed
    bTruncated       : BOOL;                  // 超目标长度发生截断 / truncation to the target length happened
END_VAR
VAR CONSTANT
    DL_STR_CAP_MAX   : USINT := 255;          // STRING 型长度上限 [字符]，R49 口径 / STRING capacity [characters], per R49
    DL_STR_TARGET_MIN : USINT := 1;           // 目标长度下限 [字符] / target length lower bound [characters]
    DL_STR_SCAN_MAX  : INT := 255;            // 扫描上界 [字符]，与 STRING 上限一致 / scan bound [characters], equals the STRING capacity
    DL_STR_BLANK     : STRING(1) := ' ';      // 单个空格字符，修剪判据 / a single blank used by the trim test
    DL_STR_EMPTY     : STRING(1) := '';       // 空串常量，故障缺省返回 / empty string returned on faults
    DL_STR_NAN       : STRING(3) := 'NaN';    // 统一 NaN 文本 / the unified NaN text
    DL_STR_INF_POS   : STRING(4) := 'Inf+';   // 统一正无穷文本 / the unified positive infinity text
    DL_STR_INF_NEG   : STRING(4) := 'Inf-';   // 统一负无穷文本 / the unified negative infinity text
    DL_LREAL_INF_ABS : LREAL := 1.7976931348623157E308; // 无穷幅值兜底阈值＝LREAL 最大值 [无量纲] / fallback magnitude threshold equal to the LREAL maximum [dimensionless]
    DL_LREAL_ZERO    : LREAL := 0.0;          // 浮点零常量，符号判定用 [无量纲] / float zero constant used by the sign test [dimensionless]
    DL_INT_ZERO      : INT := 0;              // 整型零常量，避免裸字面量 [字符] / integer zero constant [characters]
    DL_INT_ONE       : INT := 1;              // 整型一常量，首个非空格位置起点 [字符] / integer one constant, first non-blank position [characters]
END_VAR
VAR
    sText            : STRING(255);           // 文本中间串，有限与非有限共用 / text intermediate shared by both branches
    sTrim            : STRING(255);           // 修剪后的中间串 / intermediate string after the trim
    sOut             : STRING(255);           // 最终输出串 / final output string
    sChar            : STRING(1);             // 单字符比较缓冲 / single character comparison buffer
    nLen             : INT;                   // 中间串有效长度 [字符] / effective length of the intermediate string [characters]
    nStart           : INT;                   // 首个非空格位置，1 起始，0 = 全为空格 / first non-blank position, 1-based, 0 means all blanks
    nIdx             : INT;                   // 扫描游标 [字符]，1 起始 / scan cursor [characters], 1-based
    nKept            : INT;                   // 修剪后保留长度，一次锁存 [字符] / retained length, latched exactly once [characters]
    nTarget          : INT;                   // 目标长度，由引脚转出并钳位 [字符] / target length derived and clamped [characters]
    bFound           : BOOL;                  // 已找到首个非空格标志 / a first non-blank has been found
    bNaN             : BOOL;                  // 自反性判据命中的 NaN 标志 / NaN hit by the reflexivity test
    bInf             : BOOL;                  // 幅值判据命中的无穷标志 / infinity hit by the magnitude test
END_VAR

// 段 1｜返回值与错误状态预置 / segment 1, preset return value and error status
FC_DL_LrealToStringTrim := DL_STR_EMPTY;      // 故障缺省返回空串 / fault default returns an empty string
eErr := 0;                                    // 预置无错误 / preset no error
bError := FALSE;                              // 预置无故障 / preset no fault
bValid := FALSE;                              // 预置不可用，通过闸门后置位 / preset invalid, set TRUE after the gates
bNonFinite := FALSE;                          // 预置有限输入 / preset finite input
bTrimmed := FALSE;                            // 预置未修剪 / preset no trim
bTruncated := FALSE;                          // 预置未截断 / preset no truncation
sText := DL_STR_EMPTY;                        // 文本中间串清零 / clear the text intermediate
nKept := DL_INT_ZERO;                         // 保留长度清零 / clear the retained length

// 段 2｜目标长度钳位（0 长度无意义，结构性钳到 1，钳位后果由截断分支显式体现）/ segment 2, target length clamp
nTarget := USINT_TO_INT(uTargetMax);          // 目标长度转整型 [字符] / convert the target length into an integer [characters]
IF nTarget < USINT_TO_INT(DL_STR_TARGET_MIN) THEN
    nTarget := USINT_TO_INT(DL_STR_TARGET_MIN); // 0 长度目标钳到 1 字符 / a zero target is clamped to one character
END_IF
IF nTarget > USINT_TO_INT(DL_STR_CAP_MAX) THEN
    nTarget := USINT_TO_INT(DL_STR_CAP_MAX);  // 双保险：按 STRING 上限钳位 [字符] / second line of defence, clamp to the STRING capacity [characters]
END_IF

// 段 3｜非有限防御闸：先判 NaN 再判无穷，两判据分开置位 / segment 3, non-finite gate with two separate tests
bNaN := fIn <> fIn;                           // IEEE 754 自反性判据：NaN 与自身比较恒假 / reflexivity test, NaN never equals itself
bInf := FALSE;                                // 无穷标志预置 / preset the infinity flag
IF NOT bNaN THEN
    bInf := ((fIn - fIn) <> (fIn - fIn)) OR (ABS(fIn) >= DL_LREAL_INF_ABS); // 双判据：x−x 在无穷处产 NaN（精确判据），幅值兜底只余「恰为最大值」单值残余 [无量纲] / dual test, x minus x yields NaN at infinity while the magnitude fallback only leaves the exact-maximum residue [dimensionless]
END_IF

IF bNaN THEN
    sText := DL_STR_NAN;                      // 统一 NaN 文本，不做内建转换 / unified NaN text, no built-in conversion
    bNonFinite := TRUE;                       // 标记非有限输入 / flag the non-finite input
    eErr := 16#0001_0428;                     // 信息级：非有限值已映射统一文本 / info level, mapped onto the unified text
ELSIF bInf THEN
    IF fIn > DL_LREAL_ZERO THEN
        sText := DL_STR_INF_POS;              // 统一正无穷文本 / unified positive infinity text
    ELSE
        sText := DL_STR_INF_NEG;              // 统一负无穷文本 / unified negative infinity text
    END_IF
    bNonFinite := TRUE;                       // 标记非有限输入 / flag the non-finite input
    eErr := 16#0001_0428;                     // 信息级：非有限值已映射统一文本 / info level, mapped onto the unified text
ELSE
    // 段 4｜有限值：委托平台内建字符串化 / segment 4, finite values go through the built-in
    sText := LREAL_TO_STRING(fIn);            // 数值 → 原始串（可能含前导空格）/ value to raw string, possibly blank padded
END_IF

// 段 5｜有效长度一次锁存并钳位 / segment 5, latch the effective length once and clamp it
nLen := LEN(sText);                           // 中间串长度 [字符] / intermediate string length [characters]
IF nLen > DL_STR_SCAN_MAX THEN
    nLen := DL_STR_SCAN_MAX;                  // 超容量按上限钳位 [字符] / clamp to the capacity [characters]
ELSIF nLen < DL_INT_ZERO THEN
    nLen := DL_INT_ZERO;                      // 负长度防御，结构性不可达 [字符] / negative length guard, structurally unreachable [characters]
END_IF

// 段 6｜前导空格修剪：定长 FOR 扫描，禁 WHILE / segment 6, leading blank trim with a bounded FOR loop
nStart := DL_INT_ZERO;                        // 0 表示尚未找到非空格 / zero means no non-blank found yet
bFound := FALSE;                              // 扫描标志预置 / preset the scan flag
FOR nIdx := DL_INT_ONE TO nLen DO
    IF NOT bFound THEN
        sChar := MID(sText, DL_INT_ONE, nIdx); // 取当前字符 / take the current character
        IF sChar <> DL_STR_BLANK THEN
            nStart := nIdx;                   // 记录首个非空格位置 [字符] / record the first non-blank position [characters]
            bFound := TRUE;                   // 扫描标志置位 / raise the scan flag
        END_IF
    END_IF
END_FOR

IF nStart = DL_INT_ZERO THEN
    sTrim := DL_STR_EMPTY;                    // 全为空格：合法的空结果，不是错误 / all blanks, a legal empty result
ELSE
    sTrim := MID(sText, nLen - nStart + DL_INT_ONE, nStart); // 一次截取中间段 / extract the retained segment in one call
    IF nStart > DL_INT_ONE THEN
        bTrimmed := TRUE;                     // 确实修剪了前导空格 / blanks were really trimmed
        eErr := 16#0001_0429;                 // 信息级：发生空格修剪 / info level, blanks were trimmed
    END_IF
END_IF

// 段 7｜四步截断样板（R37）：长度锁存 → 宽度比较 → 标志先置 → 按允许分路 / segment 7, the four-step truncation pattern
nKept := LEN(sTrim);                          // 修剪后长度，一次锁存 [字符] / retained length, latched once [characters]
IF nKept > nTarget THEN
    bTruncated := TRUE;                       // 标志先于任何写入 / the flag precedes every write
    IF bAllowTrunc THEN
        sOut := LEFT(sTrim, nTarget);         // 允许截断：按目标长度截取 / truncation allowed, take the target length
        eErr := 16#0001_0429;                 // 信息级：发生截断，值可用 / info level, truncated, still usable
    ELSE
        eErr := 16#0001_035A;                 // 故障级：需截断但不允许 / fault level, truncation needed but not allowed
        bError := TRUE;                       // 置故障标志 / raise the error flag
        bValid := FALSE;                      // 返回值不可用 / flag the return as unusable
        FC_DL_LrealToStringTrim := DL_STR_EMPTY; // 返回空串，绝不返回半截数值 / return an empty string, never a partial number
        RETURN;                               // 出口 / exit
    END_IF
ELSE
    sOut := sTrim;                            // 无需截断，直接采用修剪结果 / no truncation, take the trimmed string
END_IF

// 段 8｜发布结果 / segment 8, publish the result
FC_DL_LrealToStringTrim := sOut;              // 输出最终串 / publish the final string
bValid := TRUE;                               // 有限值与非有限统一文本均可用 / both finite and unified non-finite texts are usable
bError := FALSE;                              // 信息级不置故障（双保险）/ info level never raises a fault, second line of defence
END_FUNCTION

(* ---- FC_DL_LwordBitCount.st ---- *)
(*
    组件名称 : FC_DL_LwordBitCount
    所属子库 : DL_MathData
    当前版本 : 1.0.0
    兼 容 性 : CODESYS V3.5+ / TwinCAT 3 / 汇川 InoProShop；仅依赖 Standard.library
    功能描述 : LWORD 汉明重量（置位个数 0~64），补齐存量 FC_DL_BitCount 只覆盖 DWORD 的位宽缺口。
              取舍 ①：Brian Kernighan 法 —— 每次 u AND (u − 1) 消掉最低的一个 1，迭代次数恰等于置位数；
              全零输入零次迭代。禁改成 FOR 0..63 的定长 64 次：定长版在「稀疏字」（如只有第 63 位为 1）
              上要多做 63 次无用循环，且与库内 BitCount 的算法选择必须同源，否则两件的行为一致性无从对照。
              取舍 ②：WHILE 必带守卫计数器 —— 理论上 Kernighan 法对 64 位字最多 64 次即归零，
              守卫超限只可能是实现回归或平台整数语义异常，属必须显式落码的防御分支。
              取舍 ③：全零输入是合法工况（未接线的状态字、刚清零的报警位图），返回 0 并发信息码，
              绝不判故障 —— 把「正常空值」当故障会让诊断日志被无效条目淹没。
    开源溯源 : T2-1 LGF 计数与边沿子族（LGF 侧 BitCount 为 DWORD 口径，本件为 64 位域自有实现）；；本件为道莅 clean-room 防御性实现（仅借 LGF 分类事实/参数域/行为定义，零代码行与符号名复制）。
              算法为公开经典，零查表、零内存、零代码行复制，码位与分级 100% 自有。
    本文件内含 : FUNCTION FC_DL_LwordBitCount（单 POU，无配套类型）
    依 赖 : 无 DL_ 内部依赖；Standard.library: 无
    红线自检 : R1 ✓ 零全局变量与外部变量 ｜ R2 ✓ 零物理 IO 地址
              R3 ✓ 纯 IEC 61131-3 ｜ R4 ✓ WHILE 守卫计数器 + 超限置故障 + 结果域自证（≤ 64）
              R5 ✓ 全变量中英双语同行注释 ｜ R6 N/A 纯函数无顺序状态机，无 CASE 可写
              R7 N/A 无定时器、无沿检测实例 ｜ R8 ✓ 守卫上限与位宽常量化
    错误码   : 16#0001_0442 [信息级] 输入全零（合法工况），返回 0，bValid = TRUE
               16#0001_0443 [信息级] 预留禁用（不得挪用）
               16#0001_0381 [故障级] 守卫超限（理论不可达，纯防御），返回 0，bValid = FALSE
               16#0001_0382 [故障级] 预留禁用（不得挪用）
               16#0001_0383 [故障级] 预留禁用（不得挪用）
    码位总账 : 16#0001_0442 用 / 16#0001_0443 预留 ｜ 16#0001_0381 用 / 16#0001_0382 预留 / 16#0001_0383 预留
    遗留假设 : ① LWORD 在 InoProShop 早期固件上是否原生 64 位未实测；32 位降级会在编译期暴露，不静默错算。
              ② 返回值类型 USINT 的域 0~255 天然覆盖 0~64，无需额外夹域；此为类型推导，未逐平台实测。
    修订历史 :
        2026-11-16  v1.0.0  首版，R21 批次 2 入库
*)
FUNCTION FC_DL_LwordBitCount : USINT
VAR_INPUT
    uValue          : LWORD;  // 待计数的字，全 64 位有效 [位图] / word to inspect, all 64 bits are significant [bitmap]
END_VAR
VAR_OUTPUT
    eErr            : UDINT;  // 错误码，0=正常；16#0001_04XX 信息级 / 16#0001_03XX 故障级 / error id, 0=ok
    bError          : BOOL;   // 故障级标志，eErr 落 16#0001_03XX 时为 TRUE / fault flag, TRUE on fault-level eErr
    bValid          : BOOL;   // 返回值是否可用 / result usable flag
END_VAR
VAR
    uTemp           : LWORD;  // 逐位消去的工作副本 [位图] / working copy with bits cleared one by one [bitmap]
    nCount          : INT;    // 置位计数 0~64 [个] / population count, 0..64 [count]
    nGuard          : DINT;   // 守卫计数器，防 WHILE 失控 [次] / guard counter protecting the WHILE loop [count]
END_VAR
VAR CONSTANT
    DL_GUARD_MAX_BITS : DINT := 64;                      // 守卫上限，等于字宽（Kernighan 法最多 64 次）[次] / guard limit equals the word width [count]
    DL_LWORD_ONE      : LWORD := 16#0000_0000_0000_0001;  // 减一基元，用于 u AND (u − 1) [位图] / the decrement primitive for u AND (u minus one) [bitmap]
    DL_LWORD_ZERO     : LWORD := 0;                      // 零哨兵，终止条件 [位图] / zero sentinel, the termination test [bitmap]
    DL_ERR_NONE       : UDINT := 16#0000_0000;           // 无故障 / no error
END_VAR

// 段 1｜返回值与错误状态预置 / segment 1, preset the return value and the error state
FC_DL_LwordBitCount := 0;       // 故障缺省返回 0 / fault default returns zero
eErr   := DL_ERR_NONE;          // 预置无错误 / preset no error
bError := FALSE;                // 预置无故障 / preset no fault
bValid := FALSE;                // 预置结果不可用 / preset unusable
nCount := 0;                    // 计数清零 / clear the count
nGuard := 0;                    // 守卫清零 / clear the guard

// 段 2｜全零短路：全零是合法工况，返回 0 并发信息码 / segment 2, an all zero word is legal, not a fault
IF uValue = DL_LWORD_ZERO THEN
    FC_DL_LwordBitCount := 0;   // 置位数 0 / population count is zero
    eErr   := 16#0001_0442;     // 全零输入（信息级，不置 bError）/ all zero input, info level
    bValid := TRUE;             // 结果可用 / the result is usable
    RETURN;                     // 提前出口，不进循环 / early exit, never enter the loop
END_IF

// 段 3｜Kernighan 消位循环：每轮消掉最低的一个 1，WHILE 必带守卫 / segment 3, Kernighan loop with a mandatory guard
uTemp := uValue;                                        // 拷贝入参，不改输入 / copy the input, never modify it
WHILE (uTemp <> DL_LWORD_ZERO) AND (nGuard <= DL_GUARD_MAX_BITS) DO
    uTemp  := uTemp AND (uTemp - DL_LWORD_ONE);         // 消掉最低位的 1 / clear the lowest set bit
    nCount := nCount + 1;                               // 计数递增 / increment the count
    nGuard := nGuard + 1;                               // 守卫递增 / increment the guard
END_WHILE

// 段 4｜守卫复检：未归零说明循环失控，属实现回归，必须显式落码 / segment 4, the guard re-check catches a runaway loop
IF uTemp <> DL_LWORD_ZERO THEN
    FC_DL_LwordBitCount := 0;   // 不给可疑结果 / never emit a suspicious result
    eErr   := 16#0001_0381;     // 守卫超限（故障级，理论不可达）/ guard exceeded, fault level, unreachable in theory
    bError := TRUE;             // 置故障标志 / raise the fault flag
    RETURN;                     // bValid 保持 FALSE / bValid stays FALSE
END_IF

// 段 5｜出口 / segment 5, exit
FC_DL_LwordBitCount := INT_TO_USINT(nCount);   // 计数恒在 0~64，转换结构性安全 / the count stays within 0..64, so the cast is safe
bValid := TRUE;                                // 结果可用 / the result is usable
END_FUNCTION

(* ---- FC_DL_LwordBitFieldExtract.st ---- *)
(*
    组件名称 : FC_DL_LwordBitFieldExtract
    所属子库 : DL_MathData
    当前版本 : 1.0.0
    兼 容 性 : CODESYS V3.5+ / TwinCAT 3 / 汇川 InoProShop；仅依赖 Standard.library
    功能描述 : LWORD 单字位段读取（起始位 0~63，字段宽 1~64），补齐库内位操作族只覆盖 BYTE/WORD/DWORD 的缺口。
              取舍 ①：掩码构造分两条路径 —— 宽 64 直接取全一常量。因为 SHL(LWORD#1, 64) 的移位量等于容器位宽，
              在 IEC 61131-3 里属未定义行为（部分平台得 1、部分得 0、部分触发异常），绝不能靠「反正会被截断」蒙过去。
              取舍 ②：截取时先 AND 再移 —— 顺序反了（先右移再 AND）会把右侧相邻字段的位一起右移到低位，
              得到「看着像、其实串位」的脏结果；这是位域读最常见的实现错误。
              取舍 ③：读操作越界按可用宽度截断 + bTruncated —— 读无副作用，能读多少读多少并让调用方看得见；
              与写件（FC_DL_LwordBitFieldInsert）的「越界一律拒写」成对，是本轮登记的 R89 纪律。
              取舍 ④：宽域本身非法（≤0 或 >64）判故障而不截断 —— 那是参数错误而非边界擦边，
              静默截断会让「字段宽填成 100」这类配置错长期潜伏。
    开源溯源 : T2-1 LGF Bit Logic 子族（闭源文档只借「合并/拆分位域存在」这一分类事实与 Bit/Width 参数域）。；本件为道莅 clean-room 防御性实现（仅借 LGF 分类事实/参数域/行为定义，零代码行与符号名复制）。
              算法、掩码策略、截断/拒写纪律、码位与分级 100% 自有，零代码行与注释复制。
    本文件内含 : FUNCTION FC_DL_LwordBitFieldExtract（单 POU，无配套类型）
    依 赖 : 无 DL_ 内部依赖；Standard.library: 无
    红线自检 : R1 ✓ 零全局变量与外部变量 ｜ R2 ✓ 零物理 IO 地址
              R3 ✓ 纯 IEC 61131-3 ｜ R4 ✓ 起始位闸 + 宽域闸 + 移位量恒 < 64（禁 SHL(x,64)）+ 截断可观测
              R5 ✓ 全变量中英双语同行注释 ｜ R6 N/A 纯函数无顺序状态机，无 CASE 可写
              R7 N/A 无定时器、无沿检测实例 ｜ R8 ✓ 位宽与全一掩码常量化
    错误码   : 16#0001_043E [信息级] 起始位 + 宽超 64，已按可用位截断，bTruncated = TRUE，bValid = TRUE
               16#0001_043F [信息级] 预留禁用（不得挪用）
               16#0001_037B [故障级] 起始位越界（< 0 或 > 63），返回 0，bValid = FALSE
               16#0001_037C [故障级] 字段宽非法（≤ 0 或 > 64），返回 0，bValid = FALSE
               16#0001_037D [故障级] 预留禁用（不得挪用）
    码位总账 : 16#0001_043E 用 / 16#0001_043F 预留 ｜ 16#0001_037B 用 / 16#0001_037C 用 / 16#0001_037D 预留
    遗留假设 : ① LWORD 在 InoProShop 早期固件上是否原生 64 位未实测；若平台把 LWORD 降级为 32 位，
              本件的宽 64 路径与掩码常量会被编译期拒收（属编译期可见，不会静默错算）。
              ② SHL/SHR 对 LWORD 的移位量按 IEC 语义限于 [0, 63]，本件已结构性保证，未逐平台实测边界。
    修订历史 :
        2026-11-16  v1.0.0  首版，R21 批次 2 入库
*)
FUNCTION FC_DL_LwordBitFieldExtract : LWORD
VAR_INPUT
    uWord           : LWORD;  // 源字，全 64 位可读 [位图] / source word, all 64 bits readable [bitmap]
    nStartBit       : INT;    // 位段起始位，0~63，越界即拒算 [位] / field start bit, 0..63, rejected when out of range [bit]
    nWidth          : INT;    // 字段宽，1~64；超可用位时截断 [位] / field width, 1..64, truncated when it exceeds the available bits [bit]
END_VAR
VAR_OUTPUT
    eErr            : UDINT;  // 错误码，0=正常；16#0001_04XX 信息级 / 16#0001_03XX 故障级 / error id, 0=ok
    bError          : BOOL;   // 故障级标志，eErr 落 16#0001_03XX 时为 TRUE / fault flag, TRUE on fault-level eErr
    bValid          : BOOL;   // 返回值是否可用 / result usable flag
    bTruncated      : BOOL;   // 宽超可用位已截断，结果只含低位可用部分 / TRUE when the width was truncated to the available bits
END_VAR
VAR
    nEffWidth       : INT;    // 实际取用宽度，= MIN(nWidth, 64 − nStartBit) [位] / effective width, the smaller of the request and the remaining bits [bit]
    uMask           : LWORD;  // 未移位的字段掩码，低 nEffWidth 位为 1 [位图] / unshifted field mask with the low effective bits set [bitmap]
    uFieldShift     : LWORD;  // 已移到目标位置的掩码 [位图] / mask shifted into the target position [bitmap]
    uRet            : LWORD;  // 取出的字段值 [位图] / extracted field value [bitmap]
END_VAR
VAR CONSTANT
    DL_MASK64_ALL   : LWORD := 16#FFFF_FFFF_FFFF_FFFF;   // 全 64 位掩码，宽 64 时直取，规避 SHL(x, 64) [位图] / all ones mask used when the width is 64, avoiding SHL by 64 [bitmap]
    DL_MASK64_LSB   : LWORD := 16#0000_0000_0000_0001;   // 最低位常量，掩码构造的基元 [位图] / lowest bit, the primitive of the mask construction [bitmap]
    DL_LWORD_BITS   : INT := 64;                         // LWORD 位宽 [位] / width of a LWORD [bit]
    DL_BIT_MIN      : INT := 0;                          // 起始位下界 [位] / lower bound of the start bit [bit]
    DL_BIT_MAX      : INT := 63;                         // 起始位上界 [位] / upper bound of the start bit [bit]
    DL_WIDTH_MIN    : INT := 1;                          // 字段宽下界 [位] / lower bound of the field width [bit]
    DL_LWORD_ZERO   : LWORD := 0;                        // 零哨兵 [位图] / zero sentinel [bitmap]
    DL_ERR_NONE     : UDINT := 16#0000_0000;             // 无故障 / no error
END_VAR

// 段 1｜返回值与错误状态预置 / segment 1, preset the return value and the error state
FC_DL_LwordBitFieldExtract := DL_LWORD_ZERO;   // 故障缺省返回 0 / fault default returns zero
eErr       := DL_ERR_NONE;                     // 预置无错误 / preset no error
bError     := FALSE;                           // 预置无故障 / preset no fault
bValid     := FALSE;                           // 预置结果不可用 / preset unusable
bTruncated := FALSE;                           // 预置未截断 / preset not truncated

// 段 2｜起始位闸 / segment 2, start bit gate
IF (nStartBit < DL_BIT_MIN) OR (nStartBit > DL_BIT_MAX) THEN
    eErr   := 16#0001_037B;                    // 起始位越界（故障级）/ start bit out of range, fault level
    bError := TRUE;                            // 置故障标志 / raise the fault flag
    RETURN;                                    // 返回 0，bValid 保持 FALSE / return zero, bValid stays FALSE
END_IF

// 段 3｜宽域闸：宽 ≤ 0 与宽 > 64 都属参数错误，不做截断 / segment 3, width gate, a wrong width is a parameter error and is never truncated
IF (nWidth < DL_WIDTH_MIN) OR (nWidth > DL_LWORD_BITS) THEN
    eErr   := 16#0001_037C;                    // 字段宽非法（故障级）/ illegal field width, fault level
    bError := TRUE;                            // 置故障标志 / raise the fault flag
    RETURN;                                    // 返回 0，bValid 保持 FALSE / return zero, bValid stays FALSE
END_IF

// 段 4｜有效宽计算：越界按可用位截断（读操作可截断，见 R89）/ segment 4, effective width with truncation allowed for reads
nEffWidth := nWidth;                           // 先按请求宽度 / start from the requested width
IF (nStartBit + nWidth) > DL_LWORD_BITS THEN
    nEffWidth  := DL_LWORD_BITS - nStartBit;   // 只取起始位右侧剩余位 / keep only the bits right of the start bit
    bTruncated := TRUE;                        // 标记已截断 / mark the truncation
    eErr       := 16#0001_043E;                // 宽超可用位已截断（信息级，不置 bError）/ width truncated, info level
END_IF

// 段 5｜掩码构造：宽 64 走常量，其余移位量恒 < 64 / segment 5, mask construction, the shift is always below the container width
IF nEffWidth = DL_LWORD_BITS THEN
    uMask := DL_MASK64_ALL;                    // 宽 64 直取全一，禁 SHL(x, 64) / width 64 takes the all ones constant, never SHL by 64
ELSE
    uMask := SHL(DL_MASK64_LSB, nEffWidth) - DL_MASK64_LSB;   // 2^n − 1，得低 n 位全一 / two to the n minus one gives n low ones
END_IF

// 段 6｜先 AND 再右移：顺序反了会串入右侧邻位的脏数据 / segment 6, mask before shifting, the reverse order pulls in neighbouring bits
uFieldShift := SHL(uMask, nStartBit);          // 掩码移到目标位置 / move the mask to the target position
uRet        := SHR(uWord AND uFieldShift, nStartBit);   // 取段后右移归位 / extract and shift back into the low bits

// 段 7｜出口 / segment 7, exit
FC_DL_LwordBitFieldExtract := uRet;            // 输出字段值 / publish the field value
bValid := TRUE;                                // 结果可用（含截断后的结果）/ the result is usable, truncation included
END_FUNCTION

(* ---- FC_DL_LwordBitFieldInsert.st ---- *)
(*
    组件名称 : FC_DL_LwordBitFieldInsert
    所属子库 : DL_MathData
    当前版本 : 1.0.0
    兼 容 性 : CODESYS V3.5+ / TwinCAT 3 / 汇川 InoProShop；仅依赖 Standard.library
    功能描述 : LWORD 单字位段读改写（清位 → 取值 → 合成），与 FC_DL_LwordBitFieldExtract 构成读写对偶。
              取舍 ①：四步固定序不可交换 —— ① 算复位掩码 ② 清位 ③ 取值 ④ 合成。
              「先清后置」是读改写唯一安全序：若先把新值 OR 进去再清位，会把刚写进去的位一起清掉；
              若直接 OR 而不清位，旧值里为 1 的位永远抹不掉（写入 0 失效）。此纪律与库内 BitArrayInsert 同源。
              取舍 ②：越界一律拒写并返回原字 —— 写有不可逆副作用，「宁可一字不写」也不写半个字。
              这与读件的截断策略成对（R89）：读可截断、写必须拒。
              取舍 ③：字段值高位于宽外的部分只提示不静默 —— 调用方若把 16 位值写进 4 位字段，
              高位必然丢，必须让它看见，否则「写进去了但值不对」是最贵的故障形态。
              取舍 ④：bChanged 只在字值真变时为 TRUE —— 上层用它做配置写回节流，
              避免每次扫描都往 EEPROM 里刷一份没变的参数。
    开源溯源 : T2-1 LGF Bit Logic 子族，只借「合并/拆分位域存在」的分类事实与 Bit/Width 参数域；；本件为道莅 clean-room 防御性实现（仅借 LGF 分类事实/参数域/行为定义，零代码行与符号名复制）。
              清位-取值-合成顺序、拒写策略、码位与分级 100% 自有，零代码行与注释复制。
    本文件内含 : FUNCTION FC_DL_LwordBitFieldInsert（单 POU，无配套类型）
    依 赖 : 无 DL_ 内部依赖；Standard.library: 无
    红线自检 : R1 ✓ 零全局变量与外部变量 ｜ R2 ✓ 零物理 IO 地址
              R3 ✓ 纯 IEC 61131-3 ｜ R4 ✓ 起始位闸 + 宽域闸 + 越界拒写（返回原值）+ 移位量恒 < 64
              R5 ✓ 全变量中英双语同行注释 ｜ R6 N/A 纯函数无顺序状态机，无 CASE 可写
              R7 N/A 无定时器、无沿检测实例 ｜ R8 ✓ 位宽与全一掩码常量化
    错误码   : 16#0001_0440 [信息级] 字段值超宽高位已丢弃，结果照写，bValid = TRUE
               16#0001_0441 [信息级] 预留禁用（不得挪用）
               16#0001_037E [故障级] 起始位越界，返回原字，bValid = FALSE
               16#0001_037F [故障级] 字段宽非法（≤ 0 或 > 64），返回原字，bValid = FALSE
               16#0001_0380 [故障级] 起始位 + 宽 > 64，越界拒写，返回原字，bValid = FALSE
    码位总账 : 16#0001_0440 用 / 16#0001_0441 预留 ｜ 16#0001_037E 用 / 16#0001_037F 用 / 16#0001_0380 用
    遗留假设 : ① LWORD 在 InoProShop 早期固件上是否原生 64 位未实测；若降级为 32 位，宽 64 路径将被编译期拒收
              （编译期可见，不会静默错算）。
              ② 用 DEC 形式不可得，故 bChanged 由「新旧字按位不等」比较得出，比较的是整字而非字段，
              这是有意为之：整字比较能兜住「掩码算错但恰好字段相同」的实现回归。
    修订历史 :
        2026-11-16  v1.0.0  首版，R21 批次 2 入库
*)
FUNCTION FC_DL_LwordBitFieldInsert : LWORD
VAR_INPUT
    uBase           : LWORD;  // 原字，除目标字段外全部保持 [位图] / base word, every bit outside the field is preserved [bitmap]
    uField          : LWORD;  // 待写入字段值，只用低 nWidth 位 [位图] / field value to write, only the low bits are used [bitmap]
    nStartBit       : INT;    // 位段起始位，0~63 [位] / field start bit, 0..63 [bit]
    nWidth          : INT;    // 字段宽，1~64；越界即拒写 [位] / field width, 1..64, rejected when out of range [bit]
END_VAR
VAR_OUTPUT
    eErr            : UDINT;  // 错误码，0=正常；16#0001_04XX 信息级 / 16#0001_03XX 故障级 / error id, 0=ok
    bError          : BOOL;   // 故障级标志，eErr 落 16#0001_03XX 时为 TRUE / fault flag, TRUE on fault-level eErr
    bValid          : BOOL;   // 返回值是否可用，FALSE 时返回的是原字 / result usable flag, FALSE means the base word is returned unchanged
    bChanged        : BOOL;   // 写出后整字与输入不同即为 TRUE，供配置写回节流 / TRUE when the resulting word differs from the input, used to throttle writes
END_VAR
VAR
    uFieldMask      : LWORD;  // 已移位的字段掩码 [位图] / shifted field mask [bitmap]
    uResetMask      : LWORD;  // 字段掩码取反，用于清位 [位图] / inverted field mask used to clear the field [bitmap]
    uTemp           : LWORD;  // 清位后的中间字 [位图] / intermediate word after clearing [bitmap]
    uVal            : LWORD;  // 截到字段宽内的待写值 [位图] / value trimmed to the field width [bitmap]
    uRet            : LWORD;  // 合成结果 [位图] / composed result [bitmap]
    uHighLost       : LWORD;  // 被丢弃的字段高位，仅用于置信息码 [位图] / discarded high bits, used only for the info code [bitmap]
    uMaskRaw        : LWORD;  // 未移位的字段掩码 [位图] / unshifted field mask [bitmap]
END_VAR
VAR CONSTANT
    DL_MASK64_ALL   : LWORD := 16#FFFF_FFFF_FFFF_FFFF;   // 全 64 位掩码，宽 64 时直取，规避 SHL(x, 64) [位图] / all ones mask for width 64 [bitmap]
    DL_MASK64_LSB   : LWORD := 16#0000_0000_0000_0001;   // 最低位常量，掩码构造基元 [位图] / lowest bit, the mask primitive [bitmap]
    DL_LWORD_BITS   : INT := 64;                         // LWORD 位宽 [位] / width of a LWORD [bit]
    DL_BIT_MIN      : INT := 0;                          // 起始位下界 [位] / lower bound of the start bit [bit]
    DL_BIT_MAX      : INT := 63;                         // 起始位上界 [位] / upper bound of the start bit [bit]
    DL_WIDTH_MIN    : INT := 1;                          // 字段宽下界 [位] / lower bound of the field width [bit]
    DL_LWORD_ZERO   : LWORD := 0;                        // 零哨兵 [位图] / zero sentinel [bitmap]
    DL_ERR_NONE     : UDINT := 16#0000_0000;             // 无故障 / no error
END_VAR

// 段 1｜返回值与错误状态预置；故障缺省返回原字（拒写的不变式）/ segment 1, preset, faults return the base word unchanged
FC_DL_LwordBitFieldInsert := uBase;             // 故障缺省返回原字 / fault default returns the base word
eErr     := DL_ERR_NONE;                        // 预置无错误 / preset no error
bError   := FALSE;                              // 预置无故障 / preset no fault
bValid   := FALSE;                              // 预置结果不可用 / preset unusable
bChanged := FALSE;                              // 预置未改动 / preset unchanged

// 段 2｜起始位闸：拒写并返回原字 / segment 2, start bit gate, refuse the write and keep the base word
IF (nStartBit < DL_BIT_MIN) OR (nStartBit > DL_BIT_MAX) THEN
    eErr   := 16#0001_037E;                     // 起始位越界（故障级）/ start bit out of range, fault level
    bError := TRUE;                             // 置故障标志 / raise the fault flag
    RETURN;                                     // 返回原字 / return the base word
END_IF

// 段 3｜宽域闸：宽 ≤ 0 或 > 64 属参数错误 / segment 3, width gate, a wrong width is a parameter error
IF (nWidth < DL_WIDTH_MIN) OR (nWidth > DL_LWORD_BITS) THEN
    eErr   := 16#0001_037F;                     // 字段宽非法（故障级）/ illegal field width, fault level
    bError := TRUE;                             // 置故障标志 / raise the fault flag
    RETURN;                                     // 返回原字 / return the base word
END_IF

// 段 4｜跨字闸：写操作越界必须拒写，「宁可一字不写」/ segment 4, cross boundary gate, a write is refused rather than truncated
IF (nStartBit + nWidth) > DL_LWORD_BITS THEN
    eErr   := 16#0001_0380;                     // 越界拒写（故障级）/ out of range write refused, fault level
    bError := TRUE;                             // 置故障标志 / raise the fault flag
    RETURN;                                     // 返回原字 / return the base word
END_IF

// 段 5｜掩码构造：宽 64 走常量，其余移位量恒 < 64 / segment 5, mask construction without any undefined shift
IF nWidth = DL_LWORD_BITS THEN
    uMaskRaw := DL_MASK64_ALL;                  // 宽 64 直取全一 / width 64 takes the all ones constant
ELSE
    uMaskRaw := SHL(DL_MASK64_LSB, nWidth) - DL_MASK64_LSB;   // 2^n − 1 / two to the n minus one
END_IF
uFieldMask := SHL(uMaskRaw, nStartBit);         // 掩码移到目标位置 / move the mask into place
uResetMask := NOT uFieldMask;                   // 复位掩码 = 字段掩码取反 / the reset mask is the inverted field mask

// 段 6｜字段高位丢弃提示（只提示，不影响写入）/ segment 6, hint about the discarded high bits, writing goes on
uHighLost := uField AND uResetMask;             // 落在字段宽之外的位 / bits that fall outside the field
IF uHighLost <> DL_LWORD_ZERO THEN
    eErr := 16#0001_0440;                       // 字段值高位已丢弃（信息级，不置 bError）/ high bits dropped, info level
END_IF

// 段 7｜四步固定序：清位 → 取值 → 合成 / segment 7, the fixed four step order, clear then set
uTemp := uBase AND uResetMask;                  // ① 清位：字段位置零，其余保持 / clear the field, keep every other bit
uVal  := uField AND uMaskRaw;                   // ② 取值：截到字段宽内 / trim the value to the field width
uRet  := uTemp OR SHL(uVal, nStartBit);         // ③ 合成：移到目标位置后或入 / ④ shift into place and OR it in

// 段 8｜改动判定与出口 / segment 8, change detection and exit
IF uRet <> uBase THEN
    bChanged := TRUE;                           // 整字真变才置位，供写回节流 / set only on a real change, used to throttle writes
END_IF
FC_DL_LwordBitFieldInsert := uRet;              // 输出合成结果 / publish the composed word
bValid := TRUE;                                 // 结果可用 / the result is usable
END_FUNCTION

(* ---- FC_DL_LwordToLintSat.st ---- *)
(*
    FC_DL_LwordToLintSat —— LWORD 到 LINT 的上饱和
    ------------------------------------------------------------------
    分类      : DL_MathData / Convert
    前缀      : FC_DL_
    版本      : 1.0.0
    溯源      : IEC 61131-3 标准语义的道莅防御性实现（LWORD 64 位无符号 → LINT 64 位有符号）；
                域内委托平台内建 LWORD_TO_LINT，本件不重实现数学内核；
                上饱和出口、无损模式复核、错误分级与码位 100% 自有；
                clean-room 重写，未复制任何闭源厂商源码，参考实现仅限 MIT/Apache 许可
    平台      : 纯 IEC 61131-3，CODESYS V3.5+ / TwinCAT 3 / InoProShop 通用
    作者      : 道莅代码库 · PLC编程专家（R20）
    ------------------------------------------------------------------
    功能说明  : 与 R19 的 FC_DL_LintToUdintSat 构成 64 位交叉域对偶：那件把有符号落无符号，
                本件把无符号大计数落有符号域。
                核心防御：① 全件比较一律在 LWORD / LINT 字面量常量之间进行，
                   禁隐式跨符号域比较——64 位跨符号域的隐式提升在部分平台走无符号路径，
                   会让 9223372036854775807 与 9223372036854775808 判等（R56 纪律）；
                ② 超域值绝不进内建：LWORD_TO_LINT 在域外是回绕行为，平台间不一致，
                   这是本件与「直接强转」的本质区别；
                ③ 上饱和置 bSatHigh 供 HMI 显示封顶；无损模式下饱和升故障级；
                ④ 域内路径零钳位、零额外比较开销。
                职责边界：有符号落无符号归 FC_DL_LintToUdintSat，64 位无符号升有符号验真归
                FC_DL_UdintToLintChk（32 位端口）；本件只管 64 位上饱和。
    编译门槛  : 主路径依赖平台内建 LWORD_TO_LINT，IEC 61131-3 标准转换函数，
                三平台标准库均提供。LWORD 字面量采用 16# 十六进制形式，
                避免十进制超长字面量在部分编译器的解析差异。
    错误码    : 16#0001_041A 超 LINT 域已饱和至 9223372036854775807——信息级，值可用
                16#0001_041B 预留禁用（信息级，不得挪用）
                16#0001_0345 调用方要求无损（bRequireLossless = TRUE）却发生饱和——故障级，bValid = FALSE
                16#0001_0346 预留（故障级，不得挪用）
                16#0001_0347 预留禁用（故障级，不得挪用）
    码位总账  : 16#0001_041A 用 / 16#0001_041B 预留 ｜ 16#0001_0345 用 / 16#0001_0346 预留 / 16#0001_0347 预留
    状态机    : R6 标注 N/A —— 本组件为纯函数无顺序状态机，无 CASE 可写，非法状态不可能出现
    采样约定  : 本件无定时器、无沿检测、无状态；单拍纯计算，结论与任务周期无关。
    修订记录  : 2026-11-16 v1.0.0 首次入库（R20）
*)
FUNCTION FC_DL_LwordToLintSat : LINT
VAR_INPUT
    uIn              : LWORD;                 // 输入值 [无量纲]，全域 0~2^64−1 / input value [dimensionless], full LWORD domain
    bRequireLossless : BOOL := FALSE;         // TRUE = 发生饱和即判故障（计量/累计场景）/ TRUE turns any saturation into a fault
END_VAR
VAR_OUTPUT
    eErr             : UDINT;                 // 错误码，0=正常 / error id, 0=ok
    bError           : BOOL;                  // 故障标志，eErr 为故障级时 TRUE / error flag, TRUE on fault-level eErr
    bValid           : BOOL;                  // 返回值是否可用（要求无损却饱和时为 FALSE）/ return usable, FALSE when saturated in lossless mode
    bSatHigh         : BOOL;                  // 上饱和发生（输入 > 9223372036854775807）/ high saturation occurred
END_VAR
VAR CONSTANT
    DL_LINT_MAX_AS_LWORD : LWORD := 16#7FFF_FFFF_FFFF_FFFF; // LINT 上限的 LWORD 形态，即 2^63−1 [无量纲] / the LINT maximum as LWORD, 2 to the 63 minus one [dimensionless]
    DL_LINT_MAX      : LINT := 9223372036854775807; // LINT 上限值 [无量纲] / the LINT maximum value [dimensionless]
    DL_LINT_ZERO     : LINT := 0;             // 有符号零常量，避免裸字面量 [无量纲] / signed zero constant [dimensionless]
END_VAR
VAR
    liOut            : LINT;                  // 结果中间量 [无量纲] / result intermediate [dimensionless]
END_VAR

// 段 1｜返回值与错误状态预置 / segment 1, preset return value and error status
FC_DL_LwordToLintSat := DL_LINT_ZERO;         // 故障缺省返回 0 [无量纲] / fault default returns zero [dimensionless]
eErr := 0;                                    // 预置无错误 / preset no error
bError := FALSE;                              // 预置无故障 / preset no fault
bValid := FALSE;                              // 预置不可用，通过闸门后置位 / preset invalid, set TRUE after the gates
bSatHigh := FALSE;                            // 预置未饱和 / preset no saturation
liOut := DL_LINT_ZERO;                        // 结果中间量清零 / clear the result intermediate

// 段 2｜上域闸：LWORD 与 LWORD 常量比较，绝不让比较隐式跨符号域 / segment 2, upper gate with LWORD constants only
IF uIn > DL_LINT_MAX_AS_LWORD THEN
    liOut := DL_LINT_MAX;                     // 上饱和至 LINT 上限 / saturate to the LINT maximum
    bSatHigh := TRUE;                         // 标记上饱和 / flag the high saturation
    eErr := 16#0001_041A;                     // 信息级：超 LINT 域已饱和 / info level, saturated beyond the LINT domain
ELSE
    // 段 3｜域内才委托内建（域外调用是回绕不一致的根源）/ segment 3, delegate only inside the domain
    liOut := LWORD_TO_LINT(uIn);              // 域内无损降位 [无量纲] / lossless narrowing inside the domain [dimensionless]
END_IF

// 段 4｜无损模式复核（要求无损却发生饱和即故障级）/ segment 4, lossless recheck
IF bRequireLossless AND bSatHigh THEN
    eErr := 16#0001_0345;                     // 故障级：要求无损却发生饱和 / fault level, saturation under the lossless requirement
    bError := TRUE;                           // 置故障标志 / raise the error flag
    bValid := FALSE;                          // 返回值不可进结算 / the value must not enter settlements
    FC_DL_LwordToLintSat := liOut;            // 仍发布钳位值供 HMI 观察 / still publish the clamped value for observation
    RETURN;                                   // 出口 / exit
END_IF

// 段 5｜发布结果 / segment 5, publish the result
FC_DL_LwordToLintSat := liOut;                // 输出 64 位有符号结果 [无量纲] / publish the signed 64-bit result [dimensionless]
bValid := TRUE;                               // 直通或钳位均可用 / usable either way
bError := FALSE;                              // 信息级不置故障 / info level never raises a fault
END_FUNCTION

(* ---- FC_DL_LwordToLrealChk.st ---- *)
(*
    FC_DL_LwordToLrealChk —— LWORD 到 LREAL 精度告警转换
    ------------------------------------------------------------------
    分类      : DL_MathData / Convert
    前缀      : FC_DL_
    版本      : 1.0.0
    溯源      : IEC 61131-3 标准语义的道莅防御性实现
                （接口语义由 IEC 61131-3 定义，内部委托平台内建 LWORD_TO_LREAL，
                  外围统一错误码 / 钳位 / 双语文档；clean-room 重写，
                  未复制任何闭源厂商源码，参考实现仅限 MIT/Apache 许可）
    平台      : 纯 IEC 61131-3，CODESYS / TwinCAT / InoProShop 通用
    作者      : 道莅代码库 · PLC编程专家（R17）
    ------------------------------------------------------------------
    功能说明  : 将 LWORD 防御性转换为 LREAL 并作为返回值输出，转换委托平台内建 LWORD_TO_LREAL；
                nIn 超过 2^53（9007199254740992，双精度浮点尾数 53 位精度极限）时，
                值照常转换输出，仅置信息级 16#0001_020E 提示低位精度损失（bError=FALSE、bValid=TRUE）；
                与 FC_DL_LintToLrealChk 的职责边界：本件源类型为无符号 64 位位串，
                LWORD 无负值分支（类型系统保证），故不需要该件的双侧比较式；
                钳位方向：无钳位（信息级仅记录，转换结果为最接近的可表值）。
    错误码    : 16#0001_020E nIn 超 2^53 精度极限，转换值低位可能失真——信息级，正常防御
                16#0001_020F 预留禁用（信息级，不得挪用）
                16#0001_0303 预留禁用（故障级，不得挪用）
                16#0001_0304 预留禁用（故障级，不得挪用）
                16#0001_0305 预留禁用（故障级，不得挪用）
    状态机    : R6 标注 N/A —— 本组件为纯函数无顺序状态机，无 CASE 可写，非法状态不可能出现，故以本节说明替代 ELSE 兜底
    修订记录  : 2026-11-16 v1.0.0 首次入库（R17）
*)
FUNCTION FC_DL_LwordToLrealChk : LREAL
VAR_INPUT
    nIn : LWORD; // 待转换 64 位无符号位串，建议域 0 ~ 16#FFFF_FFFF_FFFF_FFFF [位] / 64-bit unsigned bit string to convert, suggested domain 0 .. 16#FFFF_FFFF_FFFF_FFFF [bit]
END_VAR
VAR_OUTPUT
    eErr   : UDINT; // 错误码，0=正常 / error id, 0=ok
    bError : BOOL;  // 是否出错，eErr 非 0 时为 TRUE / error flag, TRUE when eErr is nonzero
    bValid : BOOL;  // 输出是否有效可用 / output valid flag
END_VAR
VAR CONSTANT
    DL_LW_F53_MAX : LWORD := 9007199254740992; // 双精度浮点尾数 53 位精度极限 2^53 [无量纲] / double-precision 53-bit mantissa precision limit 2^53 [dimensionless]
    DL_LREAL_ZERO : LREAL := 0.0;              // 返回值预置零（本件无故障路径，仅作预置约定） [无量纲] / preset zero, no fault path in this component [dimensionless]
END_VAR

// 段 1｜返回值与错误状态预置 / segment 1, preset return value and error status
FC_DL_LwordToLrealChk := DL_LREAL_ZERO; // 预置 0.0（本件无故障级路径，仅作预置约定） [无量纲] / preset 0.0, no fault-level path in this component [dimensionless]
eErr   := 0;     // 预置无错误 / preset no error
bError := FALSE; // 预置无故障（本件无故障级路径） / preset no fault, no fault-level path here
bValid := FALSE; // 预置输出无效，通过精度判定后置位 / preset invalid, set TRUE after the precision check

// 段 2｜53 位精度极限判定与主体转换（末段） / segment 2, 53-bit precision limit check and main conversion (final)
FC_DL_LwordToLrealChk := LWORD_TO_LREAL(nIn); // 值照常转换（委托平台内建转换语义），本件只告警不钳位 [无量纲] / convert as-is via the built-in conversion, this component warns but never clamps [dimensionless]
IF nIn > DL_LW_F53_MAX THEN // 无符号位串仅需上界单侧比较，负值分支由类型系统结构性排除 [位] / unsigned bit string only needs the upper-bound test, negative branch excluded by the type system [bit]
    eErr := 16#0001_020E; // 信息级：超 2^53 精度极限，低位可能失真，仅记录不钳位 / info level: beyond the 2^53 precision limit, low bits may lose accuracy, recorded only
ELSE
    eErr := 0;            // 精度域内无告警 / within the precision domain, no notice
END_IF
bError := FALSE; // 信息级精度告警不置故障 / info-level precision notice never raises fault
bValid := TRUE;  // 域内或精度告警输出均有效可用 / in-domain or precision-noticed output is valid
END_FUNCTION

(* ---- FC_DL_MadZScore.st ---- *)
(*==============================================================================
 * 组件名称 (Component)  : FC_DL_MadZScore
 * 所属子库 (Sublibrary) : DL_MathData
 * 当前版本 (Version)    : 1.0.0
 * 兼容性 (Platform)     : CODESYS 3.5+ / TwinCAT 3 / 汇川 InoProShop / 施耐德 Machine Expert
 *                         仅依赖 Standard.library（ABS），零厂商私有库
 * 功能描述 (Function)   : 中位数绝对偏差（MAD）稳健离群评分（纯函数 FC）。
 *                         对样本数组取中位数 → 各样本绝对偏差取中位数（MAD）
 *                         → 稳健 z 分 = (x - median) / (1.4826·MAD)，1.4826
 *                         使 MAD 一致估计正态 σ。中位数/MAD 均为次序统计量，
 *                         抗粗大误差；与 SignalStatistics/OscillationIndex
 *                         （均值域统计）分工：本件是鲁棒统计缺口。
 * 来源标签 (Origin)     : 源矩阵 T2-1 LGF Measurement ◐ 统计族待挖（R18 备注既有），自研 clean-room
 * 边界语义 (Boundary)   : ① 样本数域闸 1..32（越域/含非有限样本 → 返回
 *                         FALSE，输出哨兵 0，还原方向不饱和 R81）；
 *                         ② MAD <= eps（过半样本恒等值）→ 无尺度基准，返回
 *                         FALSE + z 哨兵 0（退化声明，R332 端点语义）；
 *                         ③ 排序用插入排序（副本数组，不改输入）；
 *                         ④ 除法仅 z 分一处，除子 MAD 已过 eps 闸，无除零。
 * 输出语义 (Fallback)   : 返回 FALSE → fMedian/fMad/fZ 哨兵 0（调用方以返回
 *                         值判有效性，非故障级）。
 * 码位     (Codes)      : 按 R297 范式零 16# 码位硬编码（纯函数无错误码）。
 * 红线自检 (Redline)    : 7 项红线已自检：R1 零全局 ✓｜R2 零物理地址 ✓｜R3 纯 IEC ✓
 *                         R4 除零（MAD eps 闸）/NaN 拒收/域闸 ✓｜R5 双语同行注释 ✓
 *                         R6 纯函数无顺序逻辑（CASE 无涉）✓｜R7 无定时器实例 ✓
 * 验收向量 (Acceptance) : V1 样本 {1,2,3,4,100}、x=3 → median=3、MAD=1、
 *                         z=0（中位数点稳健零分，均值法被 100 拖歪而本法不受）；
 *                         V2 同样本、x=100 → z=(100-3)/(1.4826·1)≈65.42
 *                         （粗大误差高分离群分）；
 *                         V3 样本 {5,5,5,5} → MAD=0 → 返回 FALSE + z 哨兵 0
 *                         （退化声明 V3 与边界②对齐）。
 * 修订历史 (Revision)   : 2026-11-20  v1.0.0  R51 首版（批 4 · 序号 20）
 *==============================================================================*)
FUNCTION FC_DL_MadZScore : BOOL        // 返回 TRUE = 评分有效（median/MAD/z 可信）/ TRUE = score valid
VAR_IN_OUT
    afSamples : ARRAY[1..32] OF LREAL;   (* 样本数组（IN_OUT 免整组拷贝，本件不写回）[工程单位] / Sample array, read-only usage *)
END_VAR
VAR_INPUT
    nCount : INT;                        (* 有效样本数，域 1..32 [点] / Valid sample count *)
    fX     : LREAL;                      (* 待评分查询值 [工程单位] / Query value *)
END_VAR
VAR_OUTPUT
    fMedian : LREAL;                     (* 样本中位数 [工程单位] / Sample median *)
    fMad    : LREAL;                     (* 绝对偏差中位数 MAD [工程单位] / Median absolute deviation *)
    fZ      : LREAL;                     (* 稳健 z 分 [-] / Robust z score *)
END_VAR
VAR
    afWork : ARRAY[1..32] OF LREAL;      (* 排序副本工作量（不改输入数组）[-] / Sort work copy *)
    afDev  : ARRAY[1..32] OF LREAL;      (* 绝对偏差工作量 [工程单位] / Deviation work *)
    i      : INT;                        (* 外层排序游标（FC 局部量允许标准名）[-] / Outer sort cursor *)
    j      : INT;                        (* 内层排序游标 [-] / Inner sort cursor *)
    nMid   : INT;                        (* 中位下标工作量 [-] / Median index work *)
    fKey   : LREAL;                      (* 插入排序关键值工作量 [-] / Insertion key work *)
    fScale : LREAL;                      (* 尺度因子 1.4826·MAD 工作量 [工程单位] / Scale factor work *)
    bFin   : BOOL;                       (* 全样本有限当拍量 [-] / All-finite flag *)
END_VAR
VAR CONSTANT
    DL_MZD_NMAX : INT := 32;             (* 样本容量上限（与数组界一致）[点] / Sample capacity *)
    DL_MZD_EPS  : LREAL := 1.0E-12;      (* MAD 判零容差 [工程单位] / MAD epsilon *)
    DL_MZD_K    : LREAL := 1.4826;       (* MAD → σ 一致性系数（公开统计常数）[-] / Consistency constant *)
END_VAR

(* —— 段 0：输出哨兵预置（还原方向不饱和，R81） —— *)
fMedian := 0.0;                          (* 中位数哨兵 / Median sentinel *)
fMad := 0.0;                             (* MAD 哨兵 / MAD sentinel *)
fZ := 0.0;                               (* z 分哨兵 / Z sentinel *)
FC_DL_MadZScore := FALSE;                (* 返回值预置无效 / Return preset invalid *)

(* —— 段 1：样本数域闸 + 非有限拒收（NaN 自反 + Inf 差判） —— *)
IF (nCount < 1) OR (nCount > DL_MZD_NMAX) THEN
    RETURN;                              (* 数越域：哨兵 + FALSE（无后处理须补，R94） / Count out of domain *)
END_IF
bFin := TRUE;                            (* 有限标志预置 / Finite flag preset *)
i := 1;                                  (* 校验游标重置（R227） / Check cursor reset *)
WHILE i <= nCount DO                     (* 逐样本非有限校验 / Per-sample finiteness *)
    IF (afSamples[i] <> afSamples[i]) OR ((afSamples[i] - afSamples[i]) <> (afSamples[i] - afSamples[i])) THEN
        bFin := FALSE;                   (* 命中非有限样本 / Non-finite hit *)
    END_IF
    i := i + 1;                          (* 游标递进 / Cursor advance *)
END_WHILE
IF NOT bFin THEN
    RETURN;                              (* 含坏样本：哨兵 + FALSE（边界①） / Bad sample: return FALSE *)
END_IF

(* —— 段 2：副本排序（插入排序，O(n²) 对 32 点可接受） —— *)
i := 1;                                  (* 副本游标重置 / Copy cursor reset *)
WHILE i <= nCount DO
    afWork[i] := afSamples[i];           (* 复制样本（不改输入，边界③） / Copy sample *)
    i := i + 1;                          (* 游标递进 / Cursor advance *)
END_WHILE
i := 2;                                  (* 插入排序外层起点 / Insertion outer start *)
WHILE i <= nCount DO
    fKey := afWork[i];                   (* 取关键值 / Take key *)
    j := i - 1;                          (* 内层起点 / Inner start *)
    WHILE (j >= 1) AND (afWork[j] > fKey) DO
        afWork[j + 1] := afWork[j];      (* 右移腾位 / Shift right *)
        j := j - 1;                      (* 游标递退 / Cursor back *)
    END_WHILE
    afWork[j + 1] := fKey;               (* 插入落位 / Insert key *)
    i := i + 1;                          (* 外层递进 / Outer advance *)
END_WHILE

(* —— 段 3：中位数（奇取中点，偶取双中均值，除子常量 2 无除零） —— *)
nMid := (nCount + 1) / 2;                (* 中位下标（INT 整除向下取整口径） / Median index *)
IF (nCount MOD 2) = 1 THEN
    fMedian := afWork[nMid];             (* 奇数样本取中点 / Odd: middle *)
ELSE
    fMedian := 0.5 * (afWork[nCount / 2] + afWork[nCount / 2 + 1]);   (* 偶数样本取双中均值 / Even: mean of two middles *)
END_IF

(* —— 段 4：绝对偏差数组及其排序（逐行自含注释，相对指代省写为 R92 禁项） —— *)
i := 1;                                  (* 偏差游标重置 / Deviation cursor reset *)
WHILE i <= nCount DO
    afDev[i] := ABS(afSamples[i] - fMedian);   (* 绝对偏差 / Absolute deviation *)
    i := i + 1;                          (* 游标递进 / Cursor advance *)
END_WHILE
i := 1;                                  (* 偏差副本入排序工作区 / Copy deviations *)
WHILE i <= nCount DO
    afWork[i] := afDev[i];               (* 复制偏差到工作区 / Copy to work *)
    i := i + 1;                          (* 游标递进 / Cursor advance *)
END_WHILE
i := 2;                                  (* 偏差排序外层起点 / Deviation sort outer *)
WHILE i <= nCount DO
    fKey := afWork[i];                   (* 取关键值 / Take key *)
    j := i - 1;                          (* 内层起点 / Inner start *)
    WHILE (j >= 1) AND (afWork[j] > fKey) DO
        afWork[j + 1] := afWork[j];      (* 右移腾位 / Shift right *)
        j := j - 1;                      (* 游标递退 / Cursor back *)
    END_WHILE
    afWork[j + 1] := fKey;               (* 插入落位 / Insert key *)
    i := i + 1;                          (* 外层递进 / Outer advance *)
END_WHILE
IF (nCount MOD 2) = 1 THEN
    fMad := afWork[nMid];                (* 奇数 MAD 取中点 / Odd MAD middle *)
ELSE
    fMad := 0.5 * (afWork[nCount / 2] + afWork[nCount / 2 + 1]);   (* 偶数 MAD 双中均值 / Even MAD mean *)
END_IF

(* —— 段 5：尺度闸与 z 分（MAD 退化端点声明，R332；除子已过 eps 闸） —— *)
fScale := DL_MZD_K * fMad;               (* 尺度因子（乘法无除零） / Scale factor *)
IF fScale <= DL_MZD_EPS THEN
    RETURN;                              (* MAD 退化：哨兵 + FALSE（边界②） / Degenerate MAD: return FALSE *)
END_IF
fZ := (fX - fMedian) / fScale;           (* 稳健 z 分（除子 fScale > eps，无除零） / Robust z *)
FC_DL_MadZScore := TRUE;                 (* 评分有效 / Valid *)
END_FUNCTION

(* ---- FC_DL_MartensiteFinishTempCalc.st ---- *)
(*
  Component : FC_DL_MartensiteFinishTempCalc
  Category  : DL_MathData
  Type      : FC
  Complexity: C1
  VERSION   : v1.0.0
  功能      : 马氏体转变点核算：按 C/Mn/Cr/Ni 含量经验式算 Ms 点，再按固定间隔算 Mf 点，负值统一钳位到 0 °C。
  开源溯源  : 道莅原创 clean-room 自研（无外部代码引用）｜License: MIT
  边界条件  : ① 各元素含量须落在 0~10 % 可表区间，越界返回哨兵 -1；
              ② Ms 经验式仅在常规合金钢成分域内可信，超出成分域只置 xInDomain = FALSE 不拒算；
              ③ Ms/Mf 负值一律钳位 0 °C（低于室温无工程意义）。
*)
FUNCTION FC_DL_MartensiteFinishTempCalc : REAL
VAR_INPUT
    fCarbonPct : REAL;   (* 含碳量 [%] Carbon content *)
    fMnPct     : REAL;   (* 锰含量 [%] Manganese content *)
    fCrPct     : REAL;   (* 铬含量 [%] Chromium content *)
    fNiPct     : REAL;   (* 镍含量 [%] Nickel content *)
END_VAR
VAR_OUTPUT
    fMsC       : REAL;   (* 马氏体开始转变温度 [°C] Martensite start temperature *)
    fMfC       : REAL;   (* 马氏体终了转变温度 [°C] Martensite finish temperature *)
    xInDomain  : BOOL;   (* 成分在经验式适用域内标志 [-] Composition in empirical domain *)
    xValid     : BOOL;   (* 计算有效性标志 [-] Calculation valid flag *)
END_VAR
VAR CONSTANT
    DL_MS_BASE : REAL := 539.0;   (* Ms 经验式常数项 [°C] Ms intercept *)
    DL_K_C     : REAL := 423.0;   (* 碳系数 [°C/%] Carbon coefficient *)
    DL_K_MN    : REAL := 30.4;    (* 锰系数 [°C/%] Manganese coefficient *)
    DL_K_CR    : REAL := 12.1;    (* 铬系数 [°C/%] Chromium coefficient *)
    DL_K_NI    : REAL := 17.7;    (* 镍系数 [°C/%] Nickel coefficient *)
    DL_MS_MF   : REAL := 215.0;   (* Ms 与 Mf 间隔 [°C] Ms-Mf interval *)
    DL_ELEM_MAX: REAL := 10.0;    (* 元素含量可表上限 [%] Element content upper bound *)
    DL_ZERO    : REAL := 0.0;     (* 零常量 [°C] Zero constant *)
END_VAR
(* 出口预置：四出口统一预置 *)
fMsC := 0.0; fMfC := 0.0; xInDomain := FALSE; xValid := FALSE;
(* 非有限拦截：自反判 NaN，自身差值判 Inf *)
IF (fCarbonPct <> fCarbonPct) OR ((fCarbonPct - fCarbonPct) <> 0.0)
   OR (fMnPct <> fMnPct) OR ((fMnPct - fMnPct) <> 0.0)
   OR (fCrPct <> fCrPct) OR ((fCrPct - fCrPct) <> 0.0)
   OR (fNiPct <> fNiPct) OR ((fNiPct - fNiPct) <> 0.0) THEN
    FC_DL_MartensiteFinishTempCalc := -1.0;   (* 哨兵 -1：输入非有限 / Sentinel -1 non-finite *)
    RETURN;
END_IF
(* 成分域闸：负含量与超上限均视为非法输入 *)
IF (fCarbonPct < DL_ZERO) OR (fMnPct < DL_ZERO) OR (fCrPct < DL_ZERO) OR (fNiPct < DL_ZERO)
   OR (fCarbonPct > DL_ELEM_MAX) OR (fMnPct > DL_ELEM_MAX)
   OR (fCrPct > DL_ELEM_MAX) OR (fNiPct > DL_ELEM_MAX) THEN
    FC_DL_MartensiteFinishTempCalc := -1.0;   (* 哨兵 -1：成分越界 / Sentinel -1 composition out of range *)
    RETURN;
END_IF
(* Ms 经验式：Ms = 539 - 423C - 30.4Mn - 12.1Cr - 17.7Ni *)
fMsC := DL_MS_BASE
        - DL_K_C  * fCarbonPct
        - DL_K_MN * fMnPct
        - DL_K_CR * fCrPct
        - DL_K_NI * fNiPct;
(* Mf 经验式：Mf = Ms - 215，负值钳位 0 °C *)
fMfC := fMsC - DL_MS_MF;
IF fMfC < DL_ZERO THEN
    fMfC := DL_ZERO;                          (* 负值钳位 [°C] / Negative clamp *)
END_IF
IF fMsC < DL_ZERO THEN
    fMsC := DL_ZERO;                          (* 负值钳位 [°C] / Negative clamp *)
END_IF
(* 适用域标注：低碳高合金组合已超出经验式拟合区间，仅标注不拒算 *)
xInDomain := (fCarbonPct >= 0.10) AND (fCarbonPct <= 0.80);
xValid := TRUE;                               (* 链路有效 / Chain valid *)
FC_DL_MartensiteFinishTempCalc := fMsC;       (* 返回 Ms 点 [°C] / Return Ms temperature *)
END_FUNCTION

(* ---- FC_DL_MaxEx.st ---- *)
(*
    FC_DL_MaxEx —— 双值取大泛型防御包装（REAL 域）
    ------------------------------------------------------------------
    分类      : DL_MathData / MinMax
    前缀      : FC_DL_
    版本      : 1.0.0
    溯源      : IEC 61131-3 标准语义的道莅防御性实现
                （内部委托平台内建函数，外围统一错误码/钳位/双语文档；
                  未复制任何闭源厂商源码，参考实现仅限 MIT/Apache 许可）
    平台      : 纯 IEC 61131-3，CODESYS / TwinCAT / InoProShop 通用
    作者      : 道莅代码库 · PLC编程专家（R16）
    ------------------------------------------------------------------
    功能说明  : 双值取大：fA > fB 时返回 fA，否则返回 fB，比较运算委托
                `>` 运算符（IEC MAX 语义），不重实现任何数学内核；
                任一输入非有限（NaN 或 ±INF）判为故障级 16#0001_02B8，
                返回 0.0 且 bValid=FALSE（非有限值参与比较语义未定义，一律拦截）；
                钳位方向：无钳位（域内值直接比较输出，异常值故障拦截）；
                ±INF 采用平台安全幅值比较判定（阈值高于 REAL 最大有限值 3.402823E38），NaN 用自不等判定；
                信息级码位全部预留禁用（本组件无信息级路径）。
    错误码    : 16#0001_02B8 任一输入非有限（NaN 或 ±INF）——故障级，返回 0.0
                16#0001_01DC 预留禁用（信息级，不得挪用）
                16#0001_01DD 预留禁用（信息级，不得挪用）
                16#0001_02B9 预留禁用（故障级，不得挪用）
                16#0001_02BA 预留禁用（故障级，不得挪用）
    状态机    : R6 标注 N/A —— 本组件为纯函数无顺序状态机，无 CASE 可写，非法状态不可能出现，故以本节说明替代 ELSE 兜底
    修订记录  : 2026-11-16 v1.0.0 首次入库（R16）
*)
FUNCTION FC_DL_MaxEx : REAL
VAR_INPUT
    fA : REAL; // 比较值 A [无量纲] / compare value A
    fB : REAL; // 比较值 B [无量纲] / compare value B
END_VAR
VAR_OUTPUT
    eErr   : UDINT; // 错误码，0=正常 / error id, 0=ok
    bError : BOOL;  // 是否出错，eErr 非 0 时为 TRUE / error flag, TRUE when eErr is nonzero
    bValid : BOOL;  // 输出是否有效可用 / output valid flag
END_VAR
VAR CONSTANT
    DL_REAL_INF_GUARD : LREAL := 4.0E38; // REAL 域 ±INF 判定阈值，高于 REAL 最大有限值 3.402823E38 [无量纲] / REAL +/-INF guard above max finite REAL 3.402823E38
END_VAR
VAR
    bBad : BOOL; // 任一输入非有限判定结果 / non-finite detection result of either input
END_VAR

// 段 1｜返回值与错误状态预置 / segment 1, preset return value and error status
FC_DL_MaxEx := 0.0; // 故障缺省返回 0 [无量纲] / fault default returns 0
eErr   := 0;     // 预置无错误 / preset no error
bError := FALSE; // 预置无故障 / preset no fault
bValid := FALSE; // 预置无效，通过防御闸后置位 / preset invalid, set TRUE after guard passes

// 段 2｜非有限防御闸 / segment 2, non-finite guard
bBad := (fA <> fA) OR (fA > DL_REAL_INF_GUARD) OR (fA < -DL_REAL_INF_GUARD)
     OR (fB <> fB) OR (fB > DL_REAL_INF_GUARD) OR (fB < -DL_REAL_INF_GUARD); // 双输入非有限判定（NaN 自不等 + 安全幅值判 ±INF） [无量纲] / both inputs non-finite check (NaN by self-inequality, +/-INF by safe magnitude)
IF bBad THEN
    FC_DL_MaxEx := 0.0;       // 故障级返回 0 [无量纲] / fault level returns 0
    eErr   := 16#0001_02B8;   // 非有限输入故障码 / non-finite input fault id
    bError := TRUE;           // 置故障标志 / set fault flag
    bValid := FALSE;          // 输出无效 / output invalid
    RETURN;                   // 立即返回 / immediate return
END_IF

// 段 3｜域内取大主体计算（末段） / segment 3, in-domain maximum main calculation (final)
IF fA > fB THEN
    FC_DL_MaxEx := fA; // A 较大，输出 A / A is larger, output A
ELSE
    FC_DL_MaxEx := fB; // B 较大或相等，输出 B（相等时二者同值） / B is larger or equal, output B (identical when equal)
END_IF
bValid := TRUE; // 域内输出有效可用 / in-domain output is valid
END_FUNCTION

(* ---- FC_DL_MaxNanEx.st ---- *)
(*
    FC_DL_MaxNanEx —— 三输入取大内建防御包装（LREAL 域）
    ------------------------------------------------------------------
    分类      : DL_MathData / MinMax
    前缀      : FC_DL_
    版本      : 1.0.0
    溯源      : IEC 61131-3 标准语义的道莅防御性实现
                （内部委托平台内建函数 MAX，外围统一错误码/钳位/双语文档；
                  未复制任何闭源厂商源码，参考实现仅限 MIT/Apache 许可）
    平台      : 纯 IEC 61131-3，CODESYS / TwinCAT / InoProShop 通用
    作者      : 道莅代码库 · PLC编程专家（R40）
    ------------------------------------------------------------------
    功能说明  : 三输入取大：返回 fA、fB、fC 中的最大值，比较内核委托平台
                内建 MAX，不重实现任何数学内核；
                四段式口径（R45①）：返回值与错误码预置安全值 → 非有限域闸命中
                不调内建直接 RETURN → 域内委托内建 MAX → 结果非有限复检兜底；
                任一输入非有限判为故障级 16#0001_03C9，返回 0.0 且 bValid=FALSE
                （NaN 参与 MAX 比较在三平台传播行为不一致，一律拦截）；
                非有限判定口径（R15）：NaN 用自不等 f <> f 判定；±Inf 用
                (f − f) <> (f − f) 差值自减判定（有限值差恒为 0，无穷处产 NaN），
                禁用近似幅值阈值——LREAL 最大有限值 1.7976931348623157E308 之上
                无可表常量，近似阈值会在近似带内制造假阳性。
    错误码    : 16#0001_03C9 任一输入非有限（NaN 或 ±Inf）——故障级，返回 0.0
    状态机    : R6 标注 N/A —— 本组件为纯函数无顺序状态机，无 CASE 可写，
                非法状态不可能出现，故以本节说明替代 ELSE 兜底
    修订记录  : 2026-11-19 v1.0.0 首次入库（R40 · 批 1 · T0 快车道）
*)
FUNCTION FC_DL_MaxNanEx : LREAL
VAR_INPUT
    fA : LREAL; // 候选值一 [无量纲] ｜ first candidate value
    fB : LREAL; // 候选值二 [无量纲] ｜ second candidate value
    fC : LREAL; // 候选值三 [无量纲] ｜ third candidate value
END_VAR
VAR_OUTPUT
    eErr   : UDINT; // 错误码，0=正常，16#0001_03XX=故障级 ｜ error id, 0=ok, 16#0001_03XX=fault level
    bError : BOOL;  // 是否出错，eErr 落故障级时为 TRUE ｜ fault flag, TRUE when eErr is fault level
    bValid : BOOL;  // 输出是否有效可用 ｜ output valid flag
END_VAR
VAR
    bBad : BOOL;  // 三输入非有限判定结果（NaN 或 ±Inf）｜ non-finite detection result of the three inputs
    fOut : LREAL; // 内建 MAX 结果暂存，供出口复检 ｜ staging of the MAX result for exit recheck
END_VAR

// 段 1｜返回值与错误状态预置 ｜ segment 1, preset return value and error status
FC_DL_MaxNanEx := 0.0; // 故障缺省返回 0 [无量纲] ｜ fault default returns 0
eErr   := 0;     // 预置无错误 ｜ preset no error
bError := FALSE; // 预置无故障 ｜ preset no fault
bValid := FALSE; // 预置无效，通过防御闸后置位 ｜ preset invalid, set TRUE after guard passes
fOut   := 0.0;   // 暂存清零 ｜ clear the staging value

// 段 2｜三输入非有限防御闸（命中不调内建，早退） ｜ segment 2, non-finite guard of the three inputs (early return, no built-in call)
bBad := (fA <> fA) OR ((fA - fA) <> (fA - fA))
     OR (fB <> fB) OR ((fB - fB) <> (fB - fB))
     OR (fC <> fC) OR ((fC - fC) <> (fC - fC)); // 三输入非有限判定：NaN 自不等 + 差值自减判 ±Inf [无量纲] ｜ non-finite check: NaN by self-inequality, +/-Inf by self-subtraction
IF bBad THEN
    FC_DL_MaxNanEx := 0.0;  // 故障级返回 0 [无量纲] ｜ fault level returns 0
    eErr   := 16#0001_03C9; // 非有限输入故障码 ｜ non-finite input fault id
    bError := TRUE;         // 置故障标志（R45 配对）｜ raise the fault flag (R45 pairing)
    bValid := FALSE;        // 输出无效 ｜ output invalid
    RETURN;                 // 早退，不调内建 ｜ early return, no built-in call
END_IF

// 段 3｜域内委托内建 MAX 内核 ｜ segment 3, delegate to the built-in MAX kernel in domain
fOut := MAX(fA, fB, fC); // 三输入取大委托内建 [无量纲] ｜ three-input maximum delegated to the built-in

// 段 4｜结果复检兜底（理论不可达：有限值的 MAX 恒有限） ｜ segment 4, exit recheck (unreachable: MAX of finite values is finite)
IF (fOut <> fOut) OR ((fOut - fOut) <> (fOut - fOut)) THEN
    FC_DL_MaxNanEx := 0.0;  // 复检失败按非有限处置 [无量纲] ｜ recheck failure treated as non-finite
    eErr   := 16#0001_03C9; // 复用非有限输入码（同因同码，不新占码位）｜ reuse the non-finite code (same cause, no new code)
    bError := TRUE;         // 置故障标志 ｜ raise the fault flag
    bValid := FALSE;        // 输出无效 ｜ output invalid
    RETURN;                 // 早退 ｜ early return
END_IF

// 段 5｜出口装配 ｜ segment 5, exit assembly
FC_DL_MaxNanEx := fOut; // 取大结果直通 ｜ maximum result pass-through
bError := FALSE;        // 正常出口不置故障 ｜ normal exit raises no fault
bValid := TRUE;         // 输出有效可用 ｜ output valid
END_FUNCTION
